(* IEC 61131-3 sources: 2026_Projet_YGO_ExcavatriceDragage/TOOLS/TEST_AUTO_CI/RESULTS/L_SIMULATION/reports (part 3) *)

(* ---- FB_Sim_PositionSensor_test.st ---- *)
(* T300 - Tests unitaires du capteur cumulatif M3. *)
TEST 'TC-T300-SEN-010 Hysteresis cumulative conserve le mot thermometre'
VAR
    fb : FB_Sim_PositionSensor;
END_VAR
    fb.Enable := TRUE;
    fb.Threshold_M := 5.0;
    fb.Hysteresis_M := 0.02;
    fb.Position_M := 4.99;
    fb();
    ASSERT_TRUE(fb.ElectricalOutput, 'Position sous seuil active DI cumulative');
    fb.Position_M := 5.01;
    fb();
    ASSERT_TRUE(fb.ElectricalOutput, 'Hysteresis maintient DI dans la bande');
    fb.Position_M := 5.03;
    fb();
    ASSERT_FALSE(fb.ElectricalOutput, 'Sortie au-dessus de seuil+hysteresis');
    fb.Position_M := 4.99;
    fb();
    ASSERT_FALSE(fb.ElectricalOutput, 'Retour dans bande ne re-declenche pas');
    fb.Position_M := 4.97;
    fb();
    ASSERT_TRUE(fb.ElectricalOutput, 'Retour sous seuil-hysteresis re-declenche');
END_TEST

TEST 'TC-T300-SEN-030 Episode intermittent est borne et rejoint la position'
VAR
    fb : FB_Sim_PositionSensor;
    i : INT;
END_VAR
    fb.Enable := TRUE;
    fb.Threshold_M := 5.0;
    fb.Position_M := 4.0;
    fb.IntermittenceActive := TRUE;
    fb.IntermittenceDurationS := 1.0;
    fb.IntermittencePeriodS := 0.12;
    fb.CycleTimeS := 0.01;
    fb();
    fb.Position_M := 6.0;
    FOR i := 1 TO 120 DO
        fb();
    END_FOR;
    ASSERT_FALSE(fb.EpisodeActive, 'Episode termine avant 1.2 s');
    ASSERT_FALSE(fb.ElectricalOutput, 'DI rejoint l etat mecanique final');
    ASSERT_GT(fb.TransitionCount, 2, 'Pertes/reprises publiees, sans front permanent');
END_TEST

TEST 'TC-T300-SEN-031 Recroisements mecaniques ne reinitialisent pas episode'
VAR
    fb : FB_Sim_PositionSensor;
    i : INT;
END_VAR
    fb.Enable := TRUE;
    fb.Threshold_M := 5.0;
    fb.Position_M := 4.0;
    fb.IntermittenceActive := TRUE;
    fb.IntermittenceDurationS := 1.0;
    fb.IntermittencePeriodS := 0.12;
    fb.CycleTimeS := 0.01;
    fb();
    FOR i := 1 TO 40 DO
        IF (i MOD 2) = 0 THEN
            fb.Position_M := 4.0;
        ELSE
            fb.Position_M := 6.0;
        END_IF;
        fb();
    END_FOR;
    fb.Position_M := 6.0;
    FOR i := 1 TO 70 DO
        fb();
    END_FOR;
    ASSERT_FALSE(fb.EpisodeActive, 'Recroisements ne prolongent pas episode au-dela de 1 s');
    ASSERT_FALSE(fb.ElectricalOutput, 'Etat final suit dernier franchissement mecanique');
END_TEST

TEST 'TC-T300-SEN-040 Cent graines deterministes bornent la stabilisation'
VAR
    fb : FB_Sim_PositionSensor;
    i : INT;
    j : INT;
END_VAR
    FOR i := 1 TO 100 DO
        fb.Enable := FALSE;
        fb();
        fb.Enable := TRUE;
        fb.Threshold_M := 5.0;
        fb.Position_M := 4.0;
        fb.IntermittenceActive := TRUE;
        fb.IntermittenceDurationS := 1.0;
        fb.IntermittencePeriodS := 0.12;
        fb.CycleTimeS := 0.01;
        fb.ScenarioSeed := DINT_TO_UDINT(i);
        fb();
        fb.Position_M := 6.0;
        FOR j := 1 TO 120 DO
            fb();
        END_FOR;
        ASSERT_FALSE(fb.EpisodeActive, 'Chaque graine termine son episode avant 1.2 s');
        ASSERT_FALSE(fb.ElectricalOutput, 'Chaque graine rejoint la position finale');
        ASSERT_GE(fb.EpisodeTogglePeriodS, 0.084, 'Periode aleatoire >= 70 % nominal');
        ASSERT_LE(fb.EpisodeTogglePeriodS, 0.156, 'Periode aleatoire <= 130 % nominal');
    END_FOR;
END_TEST

(* T300 P-A / C1-C2 — profil « BLIP COURT » : excursions electriques courtes, parametrables,
   independantes du train ~1 s ci-dessus. Signatures de la trace terrain du 2026-09-04 :
   Tremie contradictoire pendant 2 echantillons a 12,24 s ; PV reactive 1 echantillon a 14,94 s.
   Grille de test = 100 ms, celle de la trace. *)
TEST 'TC-T300-SEN-050 Blip court : largeur parametrable, deux sens, profil 1 s intact'
VAR
    fb : FB_Sim_PositionSensor;
    i : INT;
    excursions : INT;
    baseCount : UDINT;
END_VAR
    (* ---- (1) Sortie de zone, excursion 0,1 s => 1 echantillon (signature PV) ---- *)
    fb.Enable := TRUE;
    fb.Threshold_M := 5.0;
    fb.Hysteresis_M := 0.02;
    fb.CycleTimeS := 0.1;
    fb.ElectricalDelayS := 0.0;
    fb.Position_M := 4.0;
    fb();
    ASSERT_TRUE(fb.ElectricalOutput, 'Depart : dans la zone capteur');
    baseCount := fb.TransitionCount;
    fb.BlipTransitions := 1;
    fb.BlipDurationS := 0.1;
    fb.Position_M := 6.0;
    fb();
    excursions := 0;
    FOR i := 1 TO 6 DO
        fb();
        IF fb.ElectricalOutput <> fb.RawDetected THEN
            excursions := excursions + 1;
        END_IF;
    END_FOR;
    ASSERT_EQ(excursions, 1, 'Blip 0,1 s a 100 ms = 1 echantillon contradictoire');
    ASSERT_EQ(fb.TransitionCount - baseCount, 3, '1 front nominal + 2 fronts du blip');
    ASSERT_FALSE(fb.BlipActive, 'Blip borne et termine');
    ASSERT_FALSE(fb.ElectricalOutput, 'Sortie rendue a l etat mecanique final');

    (* ---- (2) Meme sens, excursion 0,2 s => 2 echantillons (signature Tremie) ---- *)
    fb.Enable := FALSE;
    fb();
    fb.Enable := TRUE;
    fb.BlipTransitions := 1;
    fb.BlipDurationS := 0.2;
    fb.Position_M := 4.0;
    fb();
    fb.Position_M := 6.0;
    fb();
    excursions := 0;
    FOR i := 1 TO 8 DO
        fb();
        IF fb.ElectricalOutput <> fb.RawDetected THEN
            excursions := excursions + 1;
        END_IF;
    END_FOR;
    ASSERT_EQ(excursions, 2, 'Blip 0,2 s a 100 ms = 2 echantillons contradictoires');
    ASSERT_FALSE(fb.ElectricalOutput, 'Sortie rendue a l etat mecanique final');

    (* ---- (3) Sens INVERSE : entree en zone (front montant) — symetrie AC5 ---- *)
    fb.Enable := FALSE;
    fb();
    fb.Enable := TRUE;
    fb.BlipTransitions := 1;
    fb.BlipDurationS := 0.2;
    fb.Position_M := 6.0;
    fb();
    ASSERT_FALSE(fb.ElectricalOutput, 'Depart : hors zone capteur');
    fb.Position_M := 4.0;
    fb();
    excursions := 0;
    FOR i := 1 TO 8 DO
        fb();
        IF fb.ElectricalOutput <> fb.RawDetected THEN
            excursions := excursions + 1;
        END_IF;
    END_FOR;
    ASSERT_EQ(excursions, 2, 'Symetrie : excursion equivalente a l entree en zone');
    ASSERT_TRUE(fb.ElectricalOutput, 'Sortie rendue a l etat mecanique final (dans la zone)');

    (* ---- (4) Blip DESACTIVE : le profil historique reste strictement inchange ---- *)
    fb.Enable := FALSE;
    fb();
    fb.Enable := TRUE;
    fb.BlipTransitions := 0;
    fb.Position_M := 4.0;
    fb();
    baseCount := fb.TransitionCount;
    fb.Position_M := 6.0;
    fb();
    excursions := 0;
    FOR i := 1 TO 10 DO
        fb();
        IF fb.ElectricalOutput <> fb.RawDetected THEN
            excursions := excursions + 1;
        END_IF;
    END_FOR;
    ASSERT_EQ(excursions, 0, 'Blip desactive : aucune excursion inventee');
    ASSERT_EQ(fb.TransitionCount - baseCount, 1, 'Blip desactive : seul le front nominal');
END_TEST

(* ---- FB_Sim_Safety_test.st ---- *)
(* =======================================================================
   Automated Unit Test - FB_Sim_Safety
   ======================================================================= *)
TEST 'TC-P13-SAF-001 Enable FALSE -> boucle AU ouverte'
VAR
    fb : FB_Sim_Safety;
END_VAR
    fb.Enable := FALSE;
    fb.SimChainOkBit := TRUE;
    fb();
    ASSERT_FALSE(fb.SimChainOk, 'Enable FALSE -> SimChainOk FALSE');
    ASSERT_FALSE(fb.SimContactorOk, 'Enable FALSE -> SimContactorOk FALSE');
END_TEST

TEST 'TC-P13-SAF-002 Pilotage boucle AU saine par SimChainOkBit et armement contacteur'
VAR
    fb : FB_Sim_Safety;
END_VAR
    fb.Enable := TRUE;
    fb.SimChainOkBit := TRUE; (* Chaine AU fermee par operateur *)
    fb();

    (* Ecoulement tempo de fermeture chaine (50ms = 60ms avancee) *)
    ADVANCE_TIME(60000000);
    fb();
    ASSERT_TRUE(fb.SimChainOk, 'SimChainOkBit TRUE -> SimChainOk TRUE apres tempo relais');

    (* Impulsion armement tenue 100ms (temps de collage contacteur) *)
    ADVANCE_TIME(10000000);
    fb.EmergencyArming := TRUE;
    fb();
    ADVANCE_TIME(110000000);
    fb();
    ASSERT_TRUE(fb.SimContactorOk, 'EmergencyArming soutenu -> SimContactorOk TRUE (engage)');

    (* Relachement impulsion -> auto-maintien *)
    ADVANCE_TIME(10000000);
    fb.EmergencyArming := FALSE;
    fb();
    ASSERT_TRUE(fb.SimContactorOk, 'Fin pulse -> Auto-maintien contacteur maintenu');
END_TEST

TEST 'TC-T306-SAF-003 Injection defaut rotation de phases par SimPhaseRotationOkBit'
VAR
    fb : FB_Sim_Safety;
END_VAR
    (* Phases saines : SimPhaseRotationOkBit=TRUE -> sortie TRUE (aucun defaut) *)
    fb.Enable := TRUE;
    fb.SimPhaseRotationOkBit := TRUE;
    fb();
    ASSERT_TRUE(fb.SimPhaseRotationOk, 'SimPhaseRotationOkBit TRUE -> SimPhaseRotationOk TRUE (phases saines)');

    (* Defaut injecte : SimPhaseRotationOkBit=FALSE -> sortie FALSE (PhaseRotationOk_DI tombe) *)
    fb.SimPhaseRotationOkBit := FALSE;
    fb();
    ASSERT_FALSE(fb.SimPhaseRotationOk, 'SimPhaseRotationOkBit FALSE -> SimPhaseRotationOk FALSE (defaut rotation de phases)');

    (* Retour a sain : nouveau passage a TRUE -> sortie TRUE *)
    fb.SimPhaseRotationOkBit := TRUE;
    fb();
    ASSERT_TRUE(fb.SimPhaseRotationOk, 'SimPhaseRotationOkBit TRUE apres FALSE -> SimPhaseRotationOk TRUE');
END_TEST

(* ---- FB_Sim_SuspendedLoad_test.st ---- *)
TEST 'TC-T300-MEC-010 Charge au repos ne cree pas d energie'
VAR
    fb : FB_Sim_SuspendedLoad;
    i : INT;
END_VAR
    fb.Enable := TRUE;
    fb.CycleTime_S := 0.01;
    FOR i := 1 TO 6000 DO
        fb();
    END_FOR;
    ASSERT_EQ(fb.Angle_Rad, 0.0, 'Angle nul sans excitation pendant 60 s');
    ASSERT_EQ(fb.AngularVelocity_RadPerS, 0.0, 'Vitesse angulaire nulle sans excitation');
END_TEST

TEST 'TC-T300-MEC-040 Acceleration excite charge et reaction reste conditionnee au frein'
VAR
    fb : FB_Sim_SuspendedLoad;
    i : INT;
END_VAR
    fb.Enable := TRUE;
    fb.CartAcceleration_Mps2 := 1.0;
    fb.BrakeMechanicallyOpen := FALSE;
    fb.CycleTime_S := 0.01;
    fb();
    ASSERT_TRUE(ABS(fb.Angle_Rad) > 0.0, 'Acceleration excite le pendule');
    ASSERT_EQ(fb.VelocityReaction_Mps, 0.0, 'Frein serre bloque reaction chariot');
    fb.BrakeMechanicallyOpen := TRUE;
    fb.CartAcceleration_Mps2 := 0.0;
    FOR i := 1 TO 10 DO
        fb();
    END_FOR;
    ASSERT_TRUE(ABS(fb.VelocityReaction_Mps) > 0.0, 'Frein ouvert publie reaction charge');
END_TEST

TEST 'TC-T300-MEC-020 Convergence pendule entre pas 10 ms et 5 ms'
VAR
    fb10 : FB_Sim_SuspendedLoad;
    fb5 : FB_Sim_SuspendedLoad;
    i : INT;
END_VAR
    fb10.Enable := TRUE;
    fb10.BrakeMechanicallyOpen := TRUE;
    fb10.CartAcceleration_Mps2 := 1.0;
    fb10.CycleTime_S := 0.01;
    fb5.Enable := TRUE;
    fb5.BrakeMechanicallyOpen := TRUE;
    fb5.CartAcceleration_Mps2 := 1.0;
    fb5.CycleTime_S := 0.005;
    fb10();
    fb5();
    fb5();
    fb10.CartAcceleration_Mps2 := 0.0;
    fb5.CartAcceleration_Mps2 := 0.0;
    FOR i := 1 TO 100 DO
        fb10();
        fb5();
        fb5();
    END_FOR;
    ASSERT_LT(ABS(fb10.Angle_Rad - fb5.Angle_Rad), 0.01,
        'Ecart angle inferieur a 10 mrad apres 1 s');
    ASSERT_LT(ABS(fb10.VelocityReaction_Mps - fb5.VelocityReaction_Mps), 0.001,
        'Ecart reaction inferieur a 1 mm/s apres 1 s');
END_TEST

(* ---- FB_Sim_Translation_test.st ---- *)
(* T300 - Tests du modele dynamique M3. *)
TEST 'TC-T300-TR-001 Etat sur desactive est P1 sans mouvement'
VAR
    fb : FB_Sim_Translation;
END_VAR
    fb.Enable := FALSE;
    fb();
    ASSERT_FALSE(fb.PosTremie, 'P1 ne doit pas annoncer Tremie');
    ASSERT_TRUE(fb.PosP1, 'Etat de repli deterministe sur P1');
    ASSERT_TRUE(fb.PosMaintenance, 'Mot thermometre P1 attendu');
    ASSERT_EQ(fb.ActualFrequency_Hz, 0.0, 'Frequence nulle');
    ASSERT_FALSE(fb.BrakeContactOpen, 'Frein ferme');
END_TEST

TEST 'TC-T300-SEN-010 Les deux extremites publient les mots thermometres valides'
VAR
    fb : FB_Sim_Translation;
    i : INT;
END_VAR
    fb.Enable := FALSE;
    fb();
    fb.Enable := TRUE;
    fb.ReqTremie := TRUE;
    fb.SpeedTgt_Pct := 100.0;
    fb.BrakeReleaseCmd := TRUE;
    fb.BrakeOpenDelayS := 0.0;
    fb.FullTravelTimeS := 0.5;
    fb.SensorElectricalDelayS := 0.0;
    FOR i := 1 TO 400 DO
        fb();
    END_FOR;
    ASSERT_TRUE(fb.PosTremie, 'Tremie active a la butee 0 m');
    ASSERT_TRUE(fb.PosPV, 'PV cumulatif actif a Tremie');
    ASSERT_TRUE(fb.PosP2, 'P2 cumulatif actif a Tremie');
    ASSERT_TRUE(fb.PosP1, 'P1 cumulatif actif a Tremie');
    ASSERT_TRUE(fb.PosMaintenance, 'Maintenance cumulatif actif a Tremie');
    ASSERT_EQ(fb.VelocityTrue_Mps, 0.0, 'Butee Tremie absorbe la vitesse chariot');

    fb.Enable := FALSE;
    fb();
    fb.Enable := TRUE;
    fb.ReqTremie := FALSE;
    fb.ReqMaintenance := TRUE;
    fb.SpeedTgt_Pct := 100.0;
    fb.BrakeReleaseCmd := TRUE;
    fb.BrakeOpenDelayS := 0.0;
    fb.FullTravelTimeS := 0.5;
    fb.SensorElectricalDelayS := 0.0;
    FOR i := 1 TO 400 DO
        fb();
    END_FOR;
    ASSERT_FALSE(fb.PosTremie, 'Tremie inactif a Maintenance');
    ASSERT_FALSE(fb.PosPV, 'PV inactif a Maintenance');
    ASSERT_FALSE(fb.PosP2, 'P2 inactif a Maintenance');
    ASSERT_FALSE(fb.PosP1, 'P1 inactif a Maintenance');
    ASSERT_FALSE(fb.PosMaintenance, 'Maintenance inactif a la butee pour mot 00000');
    ASSERT_EQ(fb.VelocityTrue_Mps, 0.0, 'Butee Maintenance absorbe la vitesse chariot');
END_TEST

TEST 'TC-T300-SEN-011 Le capteur PV commute au franchissement vers Tremie'
VAR
    fb : FB_Sim_Translation;
    i : INT;
    pvWasFalse : BOOL;
    pvTurnedTrue : BOOL;
END_VAR
    fb.Enable := TRUE;
    fb.ReqTremie := TRUE;
    fb.SpeedTgt_Pct := 100.0;
    fb.BrakeReleaseCmd := TRUE;
    fb.FullTravelTimeS := 8.0;
    fb.SensorElectricalDelayS := 0.0;
    pvWasFalse := FALSE;
    pvTurnedTrue := FALSE;
    FOR i := 1 TO 700 DO
        fb();
        IF NOT fb.PosPV THEN
            pvWasFalse := TRUE;
        END_IF;
        IF pvWasFalse AND fb.PosPV THEN
            pvTurnedTrue := TRUE;
        END_IF;
    END_FOR;
    ASSERT_TRUE(pvWasFalse, 'PV initialement inactif a P1');
    ASSERT_TRUE(pvTurnedTrue, 'PV actif apres franchissement vers Tremie');
END_TEST

TEST 'TC-T300-DRV-020 Rampe terrain 20 Hz par seconde'
VAR
    fb : FB_Sim_Translation;
    i : INT;
END_VAR
    fb.Enable := TRUE;
    fb.ReqTremie := TRUE;
    fb.SpeedTgt_Pct := 0.0;
    fb.BrakeReleaseCmd := TRUE;
    fb();
    fb.SpeedTgt_Pct := 100.0;
    FOR i := 1 TO 100 DO
        fb();
    END_FOR;
    ASSERT_GT(fb.FrequencyCmd_Hz, 19.7, 'Rampe apres 1 s >= 19.7 Hz');
    ASSERT_LT(fb.FrequencyCmd_Hz, 20.3, 'Rampe apres 1 s <= 20.3 Hz');
    ASSERT_LT(fb.ActualFrequency_Hz, fb.FrequencyCmd_Hz, 'Retour dynamique derriere la consigne');
    ASSERT_GT(fb.ActualFrequency_Hz, 16.0, 'Retour coherent avec tau 150 ms');
END_TEST

TEST 'TC-T300-BRK-025 Frein temporise et retour distinct'
VAR
    fb : FB_Sim_Translation;
    i : INT;
END_VAR
    fb.Enable := TRUE;
    fb.BrakeReleaseCmd := TRUE;
    fb.BrakeOpenDelayS := 0.10;
    fb();
    ASSERT_TRUE(fb.BrakeCoilEnergized, 'Bobine active immediatement sur ordre');
    FOR i := 1 TO 8 DO
        fb();
    END_FOR;
    ASSERT_FALSE(fb.BrakeContactOpen, 'Pas de confirmation avant 90 ms');
    fb();
    fb();
    ASSERT_TRUE(fb.BrakeMechanicallyOpen, 'Ouverture mecanique apres delai');
    ASSERT_TRUE(fb.BrakeContactOpen, 'Retour auxiliaire apres delai');
END_TEST

TEST 'TC-T300-MEC-010 Le chariot suit la frequence et excite la charge'
VAR
    fb : FB_Sim_Translation;
    i : INT;
    startPosition_M : REAL;
END_VAR
    fb.Enable := TRUE;
    fb.ReqTremie := TRUE;
    fb.SpeedTgt_Pct := 100.0;
    fb.BrakeReleaseCmd := TRUE;
    fb.BrakeOpenDelayS := 0.0;
    fb();
    startPosition_M := fb.PositionTrue_M;
    FOR i := 1 TO 100 DO
        fb();
    END_FOR;
    ASSERT_LT(fb.PositionTrue_M, startPosition_M, 'Deplacement reel vers Tremie');
    ASSERT_LT(fb.VelocityTrue_Mps, 0.0, 'Vitesse signee vers Tremie');
    ASSERT_TRUE(ABS(fb.LoadAngle_Rad) > 0.0001, 'Acceleration excite le pendule');
END_TEST

TEST 'TC-T300-MEC-030 Commandes contradictoires restent neutres'
VAR
    fb : FB_Sim_Translation;
    i : INT;
    startPosition_M : REAL;
END_VAR
    fb.Enable := TRUE;
    fb.ReqTremie := TRUE;
    fb.ReqMaintenance := TRUE;
    fb.SpeedTgt_Pct := 100.0;
    fb.BrakeReleaseCmd := TRUE;
    fb.BrakeOpenDelayS := 0.0;
    fb();
    startPosition_M := fb.PositionTrue_M;
    FOR i := 1 TO 50 DO
        fb();
    END_FOR;
    ASSERT_EQ(fb.FrequencyCmd_Hz, 0.0, 'Aucune excitation avec deux sens');
    ASSERT_EQ(fb.PositionTrue_M, startPosition_M, 'Position conservee');
END_TEST

TEST 'TC-T300-SEN-030 Episode capteur intermittent rejouable avant stabilisation'
VAR
    fb : FB_Sim_Translation;
    i : INT;
END_VAR
    fb.Enable := TRUE;
    fb.ReqMaintenance := TRUE;
    fb.SpeedTgt_Pct := 0.0;
    fb.BrakeReleaseCmd := TRUE;
    fb.BrakeOpenDelayS := 0.0;
    fb.FullTravelTimeS := 0.5;
    fb.SensorStabilizationS := 1.0;
    fb.SensorIntermittenceActive := TRUE;
    fb.SensorLoadAngleTriggerRad := 0.0;
    fb.SensorIntermittencePeriodS := 0.12;
    fb();
    fb.SpeedTgt_Pct := 100.0;
    FOR i := 1 TO 250 DO
        fb();
    END_FOR;
    ASSERT_GT(fb.SensorTransitionCount, 1, 'Au moins deux fronts DI sont publies pendant episode');
    ASSERT_FALSE(fb.PosP1, 'DI rejoint la position mecanique apres episode');
END_TEST

TEST 'TC-T300-CAM-100 Matrice 48 scenarios par 100 graines respecte invariants'
VAR
    fb : FB_Sim_Translation;
    direction : INT;
    loadProfile : INT;
    regime : INT;
    perturbation : INT;
    seed : INT;
    i : INT;
END_VAR
    FOR direction := 1 TO 2 DO
        FOR loadProfile := 1 TO 2 DO
            FOR regime := 1 TO 3 DO
                FOR perturbation := 1 TO 4 DO
                    FOR seed := 1 TO 100 DO
                        fb.Enable := FALSE;
                        fb();
                        fb.Enable := TRUE;
                        fb.ReqTremie := direction = 1;
                        fb.ReqMaintenance := direction = 2;
                        fb.SpeedTgt_Pct := 100.0;
                        fb.BrakeReleaseCmd := TRUE;
                        fb.FullTravelTimeS := 0.5;
                        fb.SensorElectricalDelayS := 0.0;
                        fb.SensorScenarioSeed := DINT_TO_UDINT(seed);
                        fb.SensorIntermittenceActive := perturbation = 3;
                        fb.SensorLoadAngleTriggerRad := 0.0;
                        IF loadProfile = 1 THEN
                            fb.LoadReactionGain_Mps2 := 0.0;
                        ELSE
                            fb.LoadReactionGain_Mps2 := 0.20;
                        END_IF;
                        IF perturbation = 4 THEN
                            fb.BrakeOpenDelayS := 0.30;
                        ELSE
                            fb.BrakeOpenDelayS := 0.0;
                        END_IF;
                        fb();
                        FOR i := 1 TO 200 DO
                            IF (regime = 2) AND (i = 80) THEN
                                fb.SpeedTgt_Pct := 0.0;
                            ELSIF (regime = 3) AND (i = 80) THEN
                                fb.SpeedTgt_Pct := 0.0;
                                fb.BrakeReleaseCmd := FALSE;
                            END_IF;
                            fb();
                            ASSERT_GE(fb.PositionTrue_M, 0.0, 'Course mecanique jamais inferieure a Tremie');
                            ASSERT_LE(fb.PositionTrue_M, 30.0, 'Course mecanique jamais superieure a Maintenance');
                            ASSERT_GE(fb.ActualFrequency_Hz, 0.0, 'Retour variateur non negatif');
                            ASSERT_LE(fb.ActualFrequency_Hz, 50.0, 'Retour variateur borne a 50 Hz');
                            IF perturbation <> 3 THEN
                                ASSERT_TRUE((NOT fb.PosTremie) OR fb.PosPV,
                                    'Mot thermometre : Tremie implique PV');
                                ASSERT_TRUE((NOT fb.PosPV) OR fb.PosP2,
                                    'Mot thermometre : PV implique P2');
                                ASSERT_TRUE((NOT fb.PosP2) OR fb.PosP1,
                                    'Mot thermometre : P2 implique P1');
                                ASSERT_TRUE((NOT fb.PosP1) OR fb.PosMaintenance,
                                    'Mot thermometre : P1 implique Maintenance');
                            END_IF;
                        END_FOR;
                    END_FOR;
                END_FOR;
            END_FOR;
        END_FOR;
    END_FOR;
END_TEST

(* T300 P-A / C4 — traversee de la faute frein dans le composite : prouve que l'entree
   descend jusqu'a FB_Sim_TranslationBrake et que la sortie remonte, sans toucher au
   nominal (premier palier d'assertions). *)
TEST 'TC-T300-BRK-041 Faute frein traverse le composite M3 (fermeture en mouvement)'
VAR
    fb : FB_Sim_Translation;
    i : INT;
END_VAR
    fb.Enable := TRUE;
    fb.ReqMaintenance := TRUE;
    fb.SpeedTgt_Pct := 100.0;
    fb.BrakeReleaseCmd := TRUE;
    fb.BrakeOpenDelayS := 0.0;
    fb();
    ASSERT_TRUE(fb.BrakeMechanicallyOpen, 'Frein ouvert au depart');
    FOR i := 1 TO 200 DO
        fb();
    END_FOR;
    ASSERT_GT(fb.ActualFrequency_Hz, 0.5, 'Chariot en mouvement (frequence non nulle)');
    ASSERT_TRUE(fb.BrakeMechanicallyOpen, 'NOMINAL : frein ouvert tant que la vitesse est non nulle');
    ASSERT_FALSE(fb.BrakeFaultCloseActive, 'Aucune faute par defaut');

    fb.BrakeFaultCloseWhileRunning := TRUE;
    FOR i := 1 TO 12 DO
        fb();
    END_FOR;
    ASSERT_TRUE(fb.BrakeFaultCloseActive, 'Faute frein relayee par le composite');
    ASSERT_GT(fb.ActualFrequency_Hz, 0.5, 'Vitesse encore non nulle a la fermeture');
    ASSERT_FALSE(fb.BrakeMechanicallyOpen, 'Faute : frein mecaniquement serre en mouvement');
END_TEST

(* T300 P-A / C3 — deceleration libre. Trace terrain 2026-09-04 : commande retiree a
   14,67 s alors que 33,98 Hz etaient retournes ; le chariot a continue d'avancer pendant
   1,49 s jusqu'a l'arret a 16,16 s. La distance de roue libre correspondante est une
   ESTIMATION (la trace ne contient aucune variable de position) : ordre de grandeur
   1,1 a 1,3 m selon la methode d'integration, jamais parcourus par le modele avant ce
   correctif qui annulait la vitesse au scan de retrait de commande.
   Le pas FullTravelTimeS est allonge (60 s) pour que le scenario reste loin des butees
   mecaniques et que l'oracle porte sur la SEULE deceleration libre, pas sur un choc. *)
TEST 'TC-T300-DRV-070 Deceleration libre : le chariot avance encore apres retrait de commande'
VAR
    fb : FB_Sim_Translation;
    i : INT;
    posAtCut_M : REAL;
END_VAR
    fb.Enable := TRUE;
    fb.ReqMaintenance := TRUE;
    fb.SpeedTgt_Pct := 100.0;
    fb.BrakeReleaseCmd := TRUE;
    fb.BrakeOpenDelayS := 0.0;
    (* Echelle par defaut du banc : palier 50 Hz (maximum variateur), 0,02 m/(Hz.s), rampe d'arret 25 Hz/s. *)
    (* Charge neutralisee : l'oracle porte sur la SEULE deceleration libre du variateur.
       Sans cela, le droop de charge (0,5 Hz par rad/s) peut faire passer ActualFrequency
       sous 39,5 Hz et rendre l'assertion de palier marginale — bruit, pas verite. *)
    fb.LoadFrequencyDroopGain_Hz := 0.0;
    fb.LoadReactionGain_Mps2 := 0.0;
    FOR i := 1 TO 400 DO
        fb();
    END_FOR;
    ASSERT_NEAR(fb.ActualFrequency_Hz, 50.0, 0.5, 'Palier 50 Hz etabli avant le retrait');
    ASSERT_LT(fb.PositionTrue_M, 30.0, 'Chariot encore hors butee (scenario non pollue)');

    (* Retrait total de la commande : plus aucune requete, consigne a zero. *)
    fb.ReqMaintenance := FALSE;
    fb.ReqTremie := FALSE;
    fb.SpeedTgt_Pct := 0.0;
    fb();
    ASSERT_GT(fb.ActualFrequency_Hz, 0.5, 'Le variateur retourne encore de la vitesse au retrait');
    posAtCut_M := fb.PositionTrue_M;

    (* Roue libre : la position doit continuer de varier tant que ActualFrequency_Hz > 0.
       Seuil = borne BASSE de la bande de reference trace (R2-O9 : 0,9 a 1,3 m). Le modele
       parcourt davantage (~2,2 m) car sa rampe de descente dure 2,0 s contre 1,49 s mesures :
       ecart de fidelite ASSUME, borne haute verifiee separement. Avant correctif : ~0,1 m. *)
    FOR i := 1 TO 300 DO
        fb();
    END_FOR;
    ASSERT_NEAR(fb.ActualFrequency_Hz, 0.0, 0.01, 'Retour variateur revenu a zero');
    ASSERT_GE(fb.PositionTrue_M - posAtCut_M, 0.9,
        'Roue libre >= borne basse trace (avant correctif : ~0,1 m)');
    ASSERT_LE(fb.PositionTrue_M - posAtCut_M, 3.0, 'Roue libre bornee (pas d emballement)');
    ASSERT_LE(fb.PositionTrue_M, 30.0, 'Course mecanique respectee');
END_TEST

(* T300 P-A / C5 — perte DEFINITIVE du capteur Tremie apres arret serre.
   Trace terrain 2026-09-04 : a 26,437 s le chariot entre en zone Tremie pendant que la
   commande est retiree ; le capteur retombe a 26,537 s et n'est JAMAIS repris sur les
   8,6 s restantes (PLAN_T300 §38 : perte unique post-arret, pas une oscillation entretenue).
   EndStopRecoilMax_M = 0 conserve le comportement historique (position ET vitesse figees,
   decision de review tracee) : les deux regimes sont verifies ici. *)
TEST 'TC-T300-SEN-052 Recul borne a la butee Tremie : DI perdue PUIS reprise oscillante (ecart trace)'
VAR
    fb : FB_Sim_Translation;
    i : INT;
    scansToFall : INT;
    scansActive : INT;
END_VAR
    (* --- (0) NON-REGRESSION : recul non autorise => comportement historique inchange --- *)
    fb.Enable := TRUE;
    fb.ReqTremie := TRUE;
    fb.SpeedTgt_Pct := 100.0;
    fb.BrakeReleaseCmd := TRUE;
    fb.BrakeOpenDelayS := 0.0;
    fb.SensorElectricalDelayS := 0.0;
    fb.EndStopRecoilMax_M := 0.0;
    (* T361 — pas de temps PINCE ici : l'oracle de ce cas est le recul a la butee, pas
       l'echelle odometrique. Le scenario vient de la trace du 2026-09-04 (quelques
       secondes de trajet) et le defaut du FB est passe de 8,0 s a 37,5 s pour s'aligner
       sur le gain reel : sans ce pas explicite, 900 scans (9 s) ne suffiraient plus a
       atteindre la butee Tremie depuis 20 m et le cas testerait autre chose que son objet. *)
    fb.FullTravelTimeS := 8.0;
    FOR i := 1 TO 900 DO
        fb();
    END_FOR;
    ASSERT_TRUE(fb.PosTremie, 'Historique : DI Tremie TENUE a la butee quand le recul est interdit');
    ASSERT_NEAR(fb.PositionTrue_M, 0.0, 0.001, 'Historique : position figee a la butee');

    (* --- (1) Recul borne autorise : la charge ressort le chariot de la zone --- *)
    fb.Enable := FALSE;
    fb();
    fb.Enable := TRUE;
    fb.EndStopRecoilMax_M := 0.5;
    fb.LoadReactionGain_Mps2 := 2.0;
    FOR i := 1 TO 900 DO
        fb();
    END_FOR;
    ASSERT_TRUE(fb.PosTremie, 'PRECONDITION : zone Tremie atteinte (recul = 0,5 m autorise)');

    (* Commande retiree a l'instant de l' entree en zone (sequence exacte de la trace). *)
    fb.ReqTremie := FALSE;
    fb.SpeedTgt_Pct := 0.0;
    scansToFall := 0;
    FOR i := 1 TO 600 DO
        fb();
        IF (NOT fb.PosTremie) AND (scansToFall = 0) THEN
            scansToFall := i;
        END_IF;
    END_FOR;
    ASSERT_GT(scansToFall, 0, 'DI Tremie RETOMBE apres l arret serre (recul borne)');
    (* Boucle a 600 scans, seuil a 300 : assertion NON tautologique, marge reelle au-dessus
       de la valeur mesuree (256 scans). *)
    ASSERT_LE(scansToFall, 300, 'Perte dans un temps borne (<= 3 s a 10 ms)');

    (* Perte DURABLE : le capteur ne se reactive pas de facon entretenue ensuite. *)
    scansActive := 0;
    FOR i := 1 TO 500 DO
        fb();
        IF fb.PosTremie THEN
            scansActive := scansActive + 1;
        END_IF;
    END_FOR;
    (* ⚠️ LIMITE CONNUE — NON MASQUEE. Le modele reduit n'a AUCUNE friction de chariot ni
       raideur de cable : le pendule amorti ramene le chariot dans la zone capteur par
       oscillations. La perte est donc BORNEE, mais pas encore DEFINITIVE comme sur la trace
       terrain (PLAN_T300 §38 : « perte unique post-arret, pas une oscillation entretenue »).
       Fermer cet ecart exige un parametre physique nouveau (friction de roulement / raideur
       de cable), hors perimetre de ce lot et non calibrable sans mesure terrain : ce test
       CARACTERISE l'etat reel, il ne le valide pas. Mesure : 106 scans actifs sur 500
       (21 %), contre 0 attendu par la trace. Assertion volontairement en enveloppe. *)
    ASSERT_LE(scansActive, 150, 'Perte BORNEE mais NON DEFINITIVE : ecart trace documente');
END_TEST

(* =========================================================================
   T361 VOLET A — ALIGNEMENT DU RATIO ODOMETRIQUE BANC / ESTIMATEUR
   =========================================================================
   Le banc et l'estimateur integrent la MEME frequence retournee, mais avec deux
   echelles construites separement :
     - estimateur (CODE/I_TRANSLATION/FB_Translation_PositionEstimator.st:153/155) :
       dx = f x GainMetersPerHzSec x dt, gain cable en PRG_05_Translation.st:591 sur
       GVL_PERSISTENT._TranslationGainMetersPerHzSec = 0,02 m/(Hz.s) (1 m/s a 50 Hz) ;
     - banc (ce FB) : dx = f x (CST_PositionAtMaintenance / (40 x FullTravelTimeS)) x dt.
   Tant que les deux echelles divergent, la position estimee prend un retard constant et
   CHAQUE franchissement de capteur produit un saut de recalage — c'est exactement ce que
   montre la trace Suivi_74 (sauts de 4,53 / 9,12 / 4,59 m, AUDIT_T360). Avec l'echelle
   historique 8,0 s le rapport valait 0,09375 / 0,02 = 4,7.
   Les deux cas ci-dessous comparent le banc a l'expression EXACTE de l'estimateur :
   ils echouent si l'une des deux echelles bouge sans l'autre. *)

TEST 'TC-T361-ALIGN-001 Ratio odometrique du banc = gain reel 0,02 m/(Hz.s)'
VAR
    fb : FB_Sim_Translation;
    i : INT;
END_VAR
    fb.Enable := TRUE;
    fb.ReqMaintenance := TRUE;
    fb.SpeedTgt_Pct := 100.0;
    fb.BrakeReleaseCmd := TRUE;
    fb.BrakeOpenDelayS := 0.0;
    (* Charge neutralisee : l'oracle porte sur l'ECHELLE seule, pas sur la reaction du pendule. *)
    fb.LoadReactionGain_Mps2 := 0.0;
    FOR i := 1 TO 400 DO
        fb();
    END_FOR;
    ASSERT_NEAR(fb.ActualFrequency_Hz, 50.0, 0.5, 'Palier 50 Hz (maximum variateur) etabli avant lecture du ratio');
    ASSERT_NEAR(fb.VelocityTrue_Mps / fb.ActualFrequency_Hz, 0.02, 0.0002,
        'Ratio banc (m/s par Hz) = _TranslationGainMetersPerHzSec (ancien : 0,09375)');
END_TEST

TEST 'TC-T361-ALIGN-002 Distance banc = integrale f x 0,02 m/(Hz.s) sur 6 s'
VAR
    fb : FB_Sim_Translation;
    i : INT;
    posStart_M : REAL;
    integralHzS : REAL;
END_VAR
    fb.Enable := TRUE;
    fb.ReqTremie := TRUE;
    fb.SpeedTgt_Pct := 100.0;
    fb.BrakeReleaseCmd := TRUE;
    fb.BrakeOpenDelayS := 0.0;
    fb.SensorElectricalDelayS := 0.0;
    fb.LoadReactionGain_Mps2 := 0.0;
    (* 2 s pour etablir le palier, puis 6 s de mesure (600 scans a 10 ms) largement
       a l'ecart des butees : 20 m -> ~15,2 m a 0,8 m/s. *)
    FOR i := 1 TO 200 DO
        fb();
    END_FOR;
    posStart_M := fb.PositionTrue_M;
    integralHzS := 0.0;
    FOR i := 1 TO 600 DO
        fb();
        integralHzS := integralHzS + fb.ActualFrequency_Hz * 0.010;
    END_FOR;
    (* Tolerance 0,25 m (soit ~5 % de 4,8 m) : elle couvre la seule trainee de 1er ordre du
       modele de vitesse, pas une erreur d'echelle — un ecart d'echelle de 4,7 ferait
       diverger les deux membres de plusieurs metres. *)
    ASSERT_NEAR(posStart_M - fb.PositionTrue_M, integralHzS * 0.02, 0.25,
        'Distance parcourue par le banc = position reconstituee par l estimateur odometrique');
END_TEST

(* Echelle de la consigne : PRG_02 envoie SpeedCmd_Pct = f / 50 Hz x 100.
   20 Hz d'approche reels = 40 % doivent redonner 20 Hz (pas 16 Hz). Charge neutralisee. *)
TEST 'TC-T417-SCALE-001 Consigne 40 pct = 20 Hz et 100 pct = 50 Hz'
VAR
    fbApproach : FB_Sim_Translation;
    fbMax : FB_Sim_Translation;
    i : INT;
END_VAR
    fbApproach.Enable := TRUE;
    fbApproach.ReqMaintenance := TRUE;
    fbApproach.SpeedTgt_Pct := 40.0;
    fbApproach.BrakeReleaseCmd := TRUE;
    fbApproach.BrakeOpenDelayS := 0.0;
    fbApproach.LoadFrequencyDroopGain_Hz := 0.0;
    fbApproach.LoadReactionGain_Mps2 := 0.0;
    fbMax.Enable := TRUE;
    fbMax.ReqMaintenance := TRUE;
    fbMax.SpeedTgt_Pct := 100.0;
    fbMax.BrakeReleaseCmd := TRUE;
    fbMax.BrakeOpenDelayS := 0.0;
    fbMax.LoadFrequencyDroopGain_Hz := 0.0;
    fbMax.LoadReactionGain_Mps2 := 0.0;
    FOR i := 1 TO 400 DO
        fbApproach();
        fbMax();
    END_FOR;
    ASSERT_NEAR(fbApproach.ActualFrequency_Hz, 20.0, 0.05, '40 pct de 50 Hz = 20 Hz en regime etabli');
    ASSERT_NEAR(fbMax.ActualFrequency_Hz, 50.0, 0.05, '100 pct = 50 Hz (maximum variateur)');
END_TEST

(* Rampe d'arret : trace reelle ~25 Hz/s (rampe variateur). Pente mesuree sur la fenetre
   utile 10 Hz -> ~4 Hz, apres le transitoire du filtre de 1er ordre. Charge neutralisee. *)
TEST 'TC-T417-DECEL-001 Pente d arret 25 Hz/s depuis l approche 20 Hz'
VAR
    fb : FB_Sim_Translation;
    i : INT;
    f1_Hz : REAL;
END_VAR
    fb.Enable := TRUE;
    fb.ReqMaintenance := TRUE;
    fb.SpeedTgt_Pct := 40.0;
    fb.BrakeReleaseCmd := TRUE;
    fb.BrakeOpenDelayS := 0.0;
    fb.LoadFrequencyDroopGain_Hz := 0.0;
    fb.LoadReactionGain_Mps2 := 0.0;
    FOR i := 1 TO 400 DO
        fb();
    END_FOR;
    ASSERT_NEAR(fb.ActualFrequency_Hz, 20.0, 0.05, 'Approche 20 Hz etablie avant le retrait');
    fb.SpeedTgt_Pct := 0.0;
    i := 0;
    WHILE (fb.ActualFrequency_Hz > 10.0) AND (i < 300) DO
        fb();
        i := i + 1;
    END_WHILE;
    f1_Hz := fb.ActualFrequency_Hz;
    FOR i := 1 TO 20 DO
        fb();
    END_FOR;
    ASSERT_NEAR((f1_Hz - fb.ActualFrequency_Hz) / 0.2, 25.0, 1.0, 'Pente de decroissance = 25 Hz/s');
END_TEST

(* Depassement apres retrait de commande a l'approche : ordre de grandeur de la trace reelle
   (~0,25 m, gain 0,02 m/(Hz.s) provisoire). Bande large : cible a confirmer par la trace 10 ms. *)
TEST 'TC-T417-OVERSHOOT-001 Depassement apres retrait a 20 Hz'
VAR
    fb : FB_Sim_Translation;
    i : INT;
    posAtCut_M : REAL;
    overshoot_M : REAL;
END_VAR
    fb.Enable := TRUE;
    fb.ReqMaintenance := TRUE;
    fb.SpeedTgt_Pct := 40.0;
    fb.BrakeReleaseCmd := TRUE;
    fb.BrakeOpenDelayS := 0.0;
    fb.LoadFrequencyDroopGain_Hz := 0.0;
    fb.LoadReactionGain_Mps2 := 0.0;
    FOR i := 1 TO 400 DO
        fb();
    END_FOR;
    ASSERT_NEAR(fb.ActualFrequency_Hz, 20.0, 0.05, 'Approche 20 Hz etablie avant le retrait');
    fb.ReqMaintenance := FALSE;
    fb.SpeedTgt_Pct := 0.0;
    fb();
    posAtCut_M := fb.PositionTrue_M;
    FOR i := 1 TO 300 DO
        fb();
    END_FOR;
    overshoot_M := fb.PositionTrue_M - posAtCut_M;
    ASSERT_GE(overshoot_M, 0.15, 'Depassement >= 0,15 m (ordre de grandeur trace reelle)');
    ASSERT_LE(overshoot_M, 0.35, 'Depassement <= 0,35 m (ordre de grandeur trace reelle)');
END_TEST

(* Acceleration du banc : chariot ET frequence retournee x facteur. L'estimateur reel integre
   f_retournee x 0,02 : il doit retrouver la distance du chariot (aucun saut de recalage). *)
TEST 'TC-SIMSPEED-001 Facteur 3 : chariot 3 m/s a 50 Hz et distance = integrale f retournee x 0,02'
VAR
    fb : FB_Sim_Translation;
    i : INT;
    posStart_M : REAL;
    integralHzS : REAL;
END_VAR
    fb.Enable := TRUE;
    fb.ReqTremie := TRUE;
    fb.SpeedTgt_Pct := 100.0;
    fb.SpeedFactor := 3.0;
    fb.BrakeReleaseCmd := TRUE;
    fb.BrakeOpenDelayS := 0.0;
    fb.SensorElectricalDelayS := 0.0;
    fb.LoadReactionGain_Mps2 := 0.0;
    FOR i := 1 TO 300 DO
        fb();
    END_FOR;
    ASSERT_NEAR(fb.ActualFrequency_Hz, 150.0, 3.0, 'frequence retournee = 3 x 50 Hz');
    ASSERT_NEAR(fb.VelocityTrue_Mps, -3.0, 0.15, 'chariot a 3 m/s (1 m/s reel x 3)');
    posStart_M := fb.PositionTrue_M;
    integralHzS := 0.0;
    FOR i := 1 TO 200 DO
        fb();
        integralHzS := integralHzS + fb.ActualFrequency_Hz * 0.010;
    END_FOR;
    ASSERT_NEAR(posStart_M - fb.PositionTrue_M, integralHzS * 0.02, 0.25,
        'estimation (f retournee x 0,02) = distance du chariot : aucun saut de recalage');
END_TEST

TEST 'TC-SIMSPEED-002 Facteur borne a 5, facteur < 1 ramene a 1'
VAR
    fb : FB_Sim_Translation;
    fbLow : FB_Sim_Translation;
    i : INT;
END_VAR
    fb.Enable := TRUE;
    fb.ReqTremie := TRUE;
    fb.SpeedTgt_Pct := 100.0;
    fb.SpeedFactor := 10.0;
    fb.BrakeReleaseCmd := TRUE;
    fb.BrakeOpenDelayS := 0.0;
    fb.LoadReactionGain_Mps2 := 0.0;
    fbLow.Enable := TRUE;
    fbLow.ReqTremie := TRUE;
    fbLow.SpeedTgt_Pct := 100.0;
    fbLow.SpeedFactor := 0.0;
    fbLow.BrakeReleaseCmd := TRUE;
    fbLow.BrakeOpenDelayS := 0.0;
    fbLow.LoadReactionGain_Mps2 := 0.0;
    FOR i := 1 TO 300 DO
        fb();
        fbLow();
    END_FOR;
    ASSERT_NEAR(fb.ActualFrequency_Hz, 250.0, 5.0, 'facteur 10 borne a 5 : 250 Hz retournes');
    ASSERT_NEAR(fbLow.ActualFrequency_Hz, 50.0, 1.0, 'facteur 0 ramene a 1 : 50 Hz retournes');
    ASSERT_NEAR(fbLow.VelocityTrue_Mps, -1.0, 0.05, 'facteur 1 : 1 m/s reel a 50 Hz');
END_TEST

(* ---- FB_Sim_TranslationBrake_test.st ---- *)
TEST 'TC-T300-BRK-010 Bobine mecanique et contact restent distincts'
VAR
    fb : FB_Sim_TranslationBrake;
    i : INT;
END_VAR
    fb.Enable := TRUE;
    fb.ReleaseCmd := TRUE;
    fb.OpenDelay_S := 0.10;
    fb.ContactDelay_S := 0.01;
    fb.CycleTime_S := 0.01;
    FOR i := 1 TO 9 DO
        fb();
    END_FOR;
    ASSERT_TRUE(fb.CoilEnergized, 'Bobine immediate');
    ASSERT_FALSE(fb.MechanicallyOpen, 'Effet mecanique pas avant delai');
    fb();
    fb();
    ASSERT_TRUE(fb.MechanicallyOpen, 'Ouverture mecanique apres 100 ms');
    fb();
    ASSERT_TRUE(fb.ContactOpen, 'Contact apres effet mecanique');
END_TEST

TEST 'TC-T300-BRK-020 Serrage attend vitesse nulle'
VAR
    fb : FB_Sim_TranslationBrake;
    i : INT;
END_VAR
    fb.Enable := TRUE;
    fb.ReleaseCmd := TRUE;
    fb.OpenDelay_S := 0.0;
    fb.CycleTime_S := 0.01;
    fb();
    fb.ReleaseCmd := FALSE;
    fb.ActualFrequency_Hz := 2.0;
    FOR i := 1 TO 20 DO
        fb();
    END_FOR;
    ASSERT_TRUE(fb.MechanicallyOpen, 'Frein reste ouvert tant que vitesse non nulle');
    fb.ActualFrequency_Hz := 0.0;
    FOR i := 1 TO 10 DO
        fb();
    END_FOR;
    ASSERT_FALSE(fb.MechanicallyOpen, 'Frein serre apres 90 ms a vitesse nulle');
END_TEST

(* T300 P-A / C4 — rejeu EXACT du defaut terrain du 2026-09-04 (trace M3, 26,437 s) :
   contact frein ferme alors que le variateur retourne encore 10,00 Hz (State.ErrorId=64).
   La branche de FAUTE est explicite et le defaut de l'entree est FALSE : le chemin nominal
   reste celui de TC-T300-BRK-020, dont la garde 0,5 Hz est validee par la MEME trace
   (frein ouvert a 0,60 Hz a 16,04 s, ferme a 0,00 Hz a 16,16 s). *)
TEST 'TC-T300-BRK-040 Faute explicite : frein M3 se ferme a 10 Hz (rejeu trace 26,437 s)'
VAR
    fb : FB_Sim_TranslationBrake;
    i : INT;
END_VAR
    fb.Enable := TRUE;
    fb.ReleaseCmd := TRUE;
    fb.OpenDelay_S := 0.0;
    fb.CloseDelay_S := 0.09;
    fb.ContactDelay_S := 0.01;
    fb.CycleTime_S := 0.01;
    fb();
    ASSERT_TRUE(fb.MechanicallyOpen, 'Frein ouvert par la commande de desserrage');
    ASSERT_FALSE(fb.FaultCloseActive, 'Faute inactive par defaut');

    (* Scenario terrain : commande retiree ET variateur retournant encore 10,00 Hz. *)
    fb.ReleaseCmd := FALSE;
    fb.ActualFrequency_Hz := 10.0;
    FOR i := 1 TO 20 DO
        fb();
    END_FOR;
    ASSERT_FALSE(fb.FaultCloseActive, 'Aucune faute injectee');
    ASSERT_TRUE(fb.MechanicallyOpen, 'NOMINAL conserve : frein OUVERT a 10,00 Hz (garde 0,5 Hz)');
    ASSERT_TRUE(fb.ContactOpen, 'NOMINAL conserve : contact toujours ouvert a 10,00 Hz');

    (* Injection explicite : fermeture hors vitesse nulle, APRES le delai de faute.
       Oracle discriminateur : si le delai de faute etait ignore, la faute serait appliquee
       des le 1er scan et l'assertion ci-dessous echouerait. *)
    fb.FaultCloseWhileRunning := TRUE;
    fb.FaultCloseDelay_S := 0.5;
    FOR i := 1 TO 4 DO
        fb();
    END_FOR;
    ASSERT_FALSE(fb.FaultCloseActive, 'Faute NON appliquee avant FaultCloseDelay_S');
    ASSERT_TRUE(fb.MechanicallyOpen, 'Frein encore ouvert pendant le delai de faute');
    FOR i := 1 TO 60 DO
        fb();
    END_FOR;
    ASSERT_TRUE(fb.FaultCloseActive, 'Branche de faute appliquee apres le delai');
    ASSERT_FALSE(fb.CoilEnergized, 'Faute : bobine retombee (etat electrique coherent)');
    ASSERT_FALSE(fb.MechanicallyOpen, 'Faute : frein MECANIQUEMENT serre a 10,00 Hz');
    ASSERT_FALSE(fb.ContactOpen, 'Faute : contact frein ferme publie a 10,00 Hz');

    (* Retrait du stimulus : retour au chemin nominal, sans etat residuel. *)
    fb.FaultCloseWhileRunning := FALSE;
    fb();
    ASSERT_FALSE(fb.FaultCloseActive, 'Retrait du stimulus : faute retombee');
END_TEST

(* ---- FB_Sim_TranslationDrive_test.st ---- *)
TEST 'TC-T300-DRV-010 Drive rampe et reponse premier ordre'
VAR
    fb : FB_Sim_TranslationDrive;
    i : INT;
END_VAR
    fb.Enable := TRUE;
    fb.FrequencyTgt_Hz := 40.0;
    fb.CycleTime_S := 0.01;
    FOR i := 1 TO 100 DO
        fb();
    END_FOR;
    ASSERT_GT(fb.FrequencyCmd_Hz, 19.7, 'Rampe 20 Hz/s apres 1 s');
    ASSERT_LT(fb.FrequencyCmd_Hz, 20.3, 'Rampe bornee apres 1 s');
    ASSERT_LT(fb.ActualFrequency_Hz, fb.FrequencyCmd_Hz, 'Retour derriere la consigne');
    ASSERT_TRUE(fb.Ready, 'Brique prete sous Enable');
END_TEST

TEST 'TC-T300-DRV-030 Charge reduit retour sans inverser la frequence'
VAR
    fb : FB_Sim_TranslationDrive;
    i : INT;
    unloaded_Hz : REAL;
END_VAR
    fb.Enable := TRUE;
    fb.FrequencyTgt_Hz := 40.0;
    fb.CycleTime_S := 0.01;
    FOR i := 1 TO 300 DO
        fb();
    END_FOR;
    unloaded_Hz := fb.ActualFrequency_Hz;
    fb.LoadAngularVelocity_RadPerS := 8.0;
    fb();
    ASSERT_LT(fb.ActualFrequency_Hz, unloaded_Hz, 'Droop charge visible au PDO');
    ASSERT_GE(fb.ActualFrequency_Hz, 0.0, 'Frequence jamais negative');
END_TEST

TEST 'TC-T300-DRV-050 Pas de 100 ms conserve le temps physique'
VAR
    fb : FB_Sim_TranslationDrive;
END_VAR
    fb.Enable := TRUE;
    fb.FrequencyTgt_Hz := 40.0;
    fb.AccelRate_HzPerS := 20.0;
    fb.CycleTime_S := 0.100;
    fb();
    ASSERT_NEAR(fb.FrequencyCmd_Hz, 2.0, 0.001,
        'A 100 ms, la rampe 20 Hz/s avance de 2 Hz');
    fb();
    ASSERT_NEAR(fb.FrequencyCmd_Hz, 4.0, 0.001,
        'Le deuxieme cycle conserve la meme duree physique');
END_TEST

(* ---- FB_SimBench_test.st ---- *)
SETUP
VAR
    FB_Bench : FB_SimBench;
    FB_SimEnc : FB_Sim_Encoder;
    FB_SimJoy : FB_Sim_Joystick;
    FB_SimSafe : FB_Sim_Safety;
    FB_SimTrans : FB_Sim_Translation;
    RawPosM1 : UDINT := 0;
    RawPosM2 : UDINT := 0;
END_VAR
END_SETUP

TEST 'TC-P03-001 Dynamique Enable : neutralisation initiale, transition Ready au repos, puis coupure'
    (* Scan 0 : Enable=FALSE -> Neutralisation *)
    FB_Bench(Enable := FALSE, RawPosM1 := RawPosM1, RawPosM2 := RawPosM2);
    ASSERT_FALSE(FB_Bench.Ready, 'Enable=FALSE -> Ready=FALSE (neutralise)');

    ADVANCE_TIME(10000000);

    (* Scan 1 : Enable=TRUE -> SimBench actif *)
    FB_Bench(Enable := TRUE, RawPosM1 := RawPosM1, RawPosM2 := RawPosM2);
    ASSERT_TRUE(FB_Bench.Ready, 'Enable=TRUE -> Ready=TRUE (nominal)');

    ADVANCE_TIME(10000000);

    (* Scan 2 : Enable=FALSE -> Re-neutralisation *)
    FB_Bench(Enable := FALSE, RawPosM1 := RawPosM1, RawPosM2 := RawPosM2);
    ASSERT_FALSE(FB_Bench.Ready, 'Coupure -> Ready retombe a FALSE');
END_TEST

TEST 'TC-P13-001 Sim_Safety : neutralisation sans Enable'
    FB_SimSafe(Enable := FALSE);
    ASSERT_FALSE(FB_SimSafe.SimChainOk, 'AU non ferme');
    ASSERT_FALSE(FB_SimSafe.SimContactorOk, 'Contacteur coupe');
END_TEST

(* =========================================================================
   AF-13 — FB_SimBench (TC-P13-010/011/012/013)
   ========================================================================= *)

TEST 'TC-P13-010 SimBench Enable=FALSE neutralise tout le banc'
    FB_Bench(Enable := FALSE, RawPosM1 := RawPosM1, RawPosM2 := RawPosM2);
    ASSERT_FALSE(FB_Bench.Ready, 'Enable=FALSE -> Ready=FALSE');
    ASSERT_FALSE(FB_Bench.Busy, 'Enable=FALSE -> Busy=FALSE');
    ASSERT_FALSE(FB_Bench.Done, 'Enable=FALSE -> Done=FALSE');
END_TEST

(* =========================================================================
   T342 — CR2 : reinjection silencieuse du comptage brut (RawPosM2 = 0 -> 1 100 000 pts)
   Remplace TC-P13-014 « initialise les codeurs absolus vierges » (ID par ailleurs porte
   par l'AF-13 pour le capteur haut TOP : collision d'ID levee au passage) : le banc
   n'initialise PLUS rien, le cas « memoire vierge » est couvert par l'initialisation
   declaree GVL_PERSISTENT._SimEncoderRawPosM1/M2 := 1000000.
   ========================================================================= *)

TEST 'TC-T342-010 AUCUNE reinjection du comptage brut : un 0 reel du codeur est conserve (pas de saut post-AU)'
    (* Etat EXACT de l'incident T338 (saut 8,50 -> 204,677 m apres reactivation du banc) :
       memoire codeur a 0, banc desactive (Enable=FALSE), puis reactivation du banc
       (GVL_Simulation.SimulationModeActive FALSE -> TRUE). Le comptage brut est un entier
       SIGNE dont le zero est arbitraire (correctif T338) : le banc ne doit JAMAIS y
       substituer une origine device, sous peine d'une teleportation de
       1 100 000 pts / 4096 pts/m = 268,55 m sur la position publiee, sans mouvement
       ni defaut, reference de homing conservee. *)
    FB_Bench(Enable := FALSE, RawPosM1 := RawPosM1, RawPosM2 := RawPosM2);
    RawPosM1 := 0;
    RawPosM2 := 0;
    ADVANCE_TIME(10000000);
    FB_Bench(Enable := TRUE, RawPosM1 := RawPosM1, RawPosM2 := RawPosM2);
    ASSERT_EQ(RawPosM2, 0, 'Reactivation : la memoire codeur M2 reste a 0 (aucune reinjection du banc)');
    ASSERT_EQ(FB_Bench.Winch.COD2_PosValue, 0, 'Aucun saut publie sur COD2_PosValue (268,55 m si reinjecte)');
    ASSERT_EQ(RawPosM1, 0, 'Reactivation : la memoire codeur M1 reste a 0 (aucune reinjection du banc)');
    ASSERT_EQ(FB_Bench.Winch.COD1_PosValue, 0, 'Aucun saut publie sur COD1_PosValue');
END_TEST

TEST 'TC-T342-011 Reactivation du banc : le comptage brut conserve sa valeur courante (aucune ecriture du banc)'
    (* Non-regression du meme invariant sur une memoire MID-COURSE (296 459 pts = la valeur
       R0 reconstituee par le diagnostic T338) : quelle que soit la valeur, la reactivation
       ne produit aucun ecart, et le banc reste sans ecriture sur la memoire du codeur. *)
    FB_Bench(Enable := FALSE, RawPosM1 := RawPosM1, RawPosM2 := RawPosM2);
    RawPosM1 := 296459;
    RawPosM2 := 296459;
    ADVANCE_TIME(10000000);
    FB_Bench(Enable := TRUE, RawPosM1 := RawPosM1, RawPosM2 := RawPosM2);
    ASSERT_EQ(RawPosM2, 296459, 'Memoire M2 mid-course inchangee par la reactivation du banc');
    ASSERT_EQ(FB_Bench.Winch.COD2_PosValue, 296459, 'Position publiee = comptage brut, sans ecart');
    ASSERT_EQ(RawPosM1, 296459, 'Memoire M1 mid-course inchangee par la reactivation du banc');
    ASSERT_EQ(FB_Bench.Winch.COD1_PosValue, 296459, 'Position publiee = comptage brut, sans ecart');
END_TEST

TEST 'TC-P13-011 SimBench 0 lecture GVL en interne (essai manuel — stub)'
    (* Stub : TC-P13-011 verifie que FB_SimBench ne lit aucune variable GVL_* en interne
       (toutes les entrees passees en parametres par PRG_02_Acquisition). Verification
       statique de code, non automatisable en boite noire. (essai manuel — stub) *)
    ASSERT_TRUE(TRUE, 'Stub : verification statique 0 lecture GVL (essai manuel)');
END_TEST

TEST 'TC-P13-012 SimBench polarite frein M1 : M1_BrakeIsOpen_DI := M1_BrakeCmd'
    FB_Bench(Enable := TRUE, M1_BrakeCmd := TRUE, RawPosM1 := RawPosM1, RawPosM2 := RawPosM2);
    ASSERT_TRUE(FB_Bench.Winch.M1_BrakeIsOpen_DI, 'M1_BrakeCmd=TRUE -> M1_BrakeIsOpen_DI=TRUE (jamais NOT)');
    ADVANCE_TIME(10000000);
    FB_Bench(Enable := TRUE, M1_BrakeCmd := FALSE, RawPosM1 := RawPosM1, RawPosM2 := RawPosM2);
    ASSERT_FALSE(FB_Bench.Winch.M1_BrakeIsOpen_DI, 'M1_BrakeCmd=FALSE -> M1_BrakeIsOpen_DI=FALSE');
END_TEST

TEST 'TC-T318-010 SimBench cable nominal independent du Kobold et injection explicite'
    FB_Bench(Enable := TRUE, SimKoboldContactValue := TRUE,
             SimM2TensionedCableFaultInject := FALSE,
             RawPosM1 := RawPosM1, RawPosM2 := RawPosM2);
    ASSERT_TRUE(FB_Bench.Winch.M2_TensionedCable_DI,
                'Kobold ne produit pas de mou de cable sans injection explicite');
    FB_Bench(Enable := TRUE, SimM2TensionedCableFaultInject := TRUE,
             RawPosM1 := RawPosM1, RawPosM2 := RawPosM2);
    ASSERT_FALSE(FB_Bench.Winch.M2_TensionedCable_DI,
                 'Injection explicite -> cable non tendu');
END_TEST

TEST 'TC-T318-020 Diagnostic electrique desactive publie etat neutre'
    FB_Bench(Enable := TRUE, SimWinchElectricalDiagnosticsActive := FALSE,
             RawPosM1 := RawPosM1, RawPosM2 := RawPosM2);
    ASSERT_EQ(FB_Bench.MotorTorqueM1_Nm, 0.0, 'Diagnostic M1 OFF -> couple neutre');
    ASSERT_FALSE(FB_Bench.MotorIsStalledM1, 'Diagnostic M1 OFF -> stall FALSE');
    ASSERT_EQ(FB_Bench.MotorTorqueM2_Nm, 0.0, 'Diagnostic M2 OFF -> couple neutre');
    ASSERT_FALSE(FB_Bench.MotorIsStalledM2, 'Diagnostic M2 OFF -> stall FALSE');
END_TEST

TEST 'TC-P13-015 SimBench delai frein M1 opt-in (T316) : SimWinchBrakeOpenDelayS retarde M1_BrakeIsOpen_DI sans jamais inverser la polarite'
    (* Delai desactive (0.0) : comportement historique, bascule au meme scan *)
    FB_Bench(Enable := TRUE, M1_BrakeCmd := TRUE, SimWinchBrakeOpenDelayS := 0.0, RawPosM1 := RawPosM1, RawPosM2 := RawPosM2);
    ASSERT_TRUE(FB_Bench.Winch.M1_BrakeIsOpen_DI, 'Delai=0.0 -> ouverture instantanee (non-regression)');
    ADVANCE_TIME(10000000);
    FB_Bench(Enable := TRUE, M1_BrakeCmd := FALSE, SimWinchBrakeOpenDelayS := 0.0, RawPosM1 := RawPosM1, RawPosM2 := RawPosM2);
    ASSERT_FALSE(FB_Bench.Winch.M1_BrakeIsOpen_DI, 'Retour delai=0.0 avant test delai>0 : etat repos');

    (* Delai actif (50 ms = 5 scans a 10 ms) : la DI reste fausse pendant le delai puis bascule *)
    ADVANCE_TIME(10000000);
    FB_Bench(Enable := TRUE, M1_BrakeCmd := TRUE, SimWinchDynamicsActive := TRUE, SimWinchBrakeOpenDelayS := 0.042, RawPosM1 := RawPosM1, RawPosM2 := RawPosM2);
    ASSERT_FALSE(FB_Bench.Winch.M1_BrakeIsOpen_DI, 'Scan 1/5 du delai : M1_BrakeIsOpen_DI reste FALSE, jamais TRUE en avance');
    ADVANCE_TIME(10000000);
    FB_Bench(Enable := TRUE, M1_BrakeCmd := TRUE, SimWinchDynamicsActive := TRUE, SimWinchBrakeOpenDelayS := 0.042, RawPosM1 := RawPosM1, RawPosM2 := RawPosM2);
    ASSERT_FALSE(FB_Bench.Winch.M1_BrakeIsOpen_DI, 'Scan 2/5 du delai : toujours FALSE');
    ADVANCE_TIME(10000000);
    FB_Bench(Enable := TRUE, M1_BrakeCmd := TRUE, SimWinchDynamicsActive := TRUE, SimWinchBrakeOpenDelayS := 0.042, RawPosM1 := RawPosM1, RawPosM2 := RawPosM2);
    ASSERT_FALSE(FB_Bench.Winch.M1_BrakeIsOpen_DI, 'Scan 3/5 du delai : toujours FALSE');
    ADVANCE_TIME(10000000);
    FB_Bench(Enable := TRUE, M1_BrakeCmd := TRUE, SimWinchDynamicsActive := TRUE, SimWinchBrakeOpenDelayS := 0.042, RawPosM1 := RawPosM1, RawPosM2 := RawPosM2);
    ASSERT_FALSE(FB_Bench.Winch.M1_BrakeIsOpen_DI, 'Scan 4/5 du delai : toujours FALSE');
    ADVANCE_TIME(10000000);
    FB_Bench(Enable := TRUE, M1_BrakeCmd := TRUE, SimWinchDynamicsActive := TRUE, SimWinchBrakeOpenDelayS := 0.042, RawPosM1 := RawPosM1, RawPosM2 := RawPosM2);
    ASSERT_TRUE(FB_Bench.Winch.M1_BrakeIsOpen_DI, 'Delai ecoule (5e scan) : M1_BrakeIsOpen_DI bascule TRUE');
END_TEST

TEST 'TC-T300-INT-010 SimBench M3 publie le retour dynamique du drive'
VAR
    i : INT;
END_VAR
    FB_Bench(Enable := TRUE, M3_ReqTremie := TRUE, M3_ReqMaintenance := FALSE,
             M3_SpeedCmd_Pct := 50.0, M3_BrakeCmd := TRUE,
             RawPosM1 := RawPosM1, RawPosM2 := RawPosM2);
    FOR i := 1 TO 20 DO
        FB_Bench(Enable := TRUE, M3_ReqTremie := TRUE, M3_ReqMaintenance := FALSE,
                 M3_SpeedCmd_Pct := 50.0, M3_BrakeCmd := TRUE,
                 RawPosM1 := RawPosM1, RawPosM2 := RawPosM2);
    END_FOR;
    ASSERT_EQ(FB_Bench.Translation.M3_StatusWord, 16#0087, 'M3 actif apres ouverture frein et retour frequence');
    FB_Bench(Enable := TRUE, M3_ReqTremie := FALSE, M3_ReqMaintenance := FALSE,
             M3_SpeedCmd_Pct := 0.0, M3_BrakeCmd := FALSE,
             RawPosM1 := RawPosM1, RawPosM2 := RawPosM2);
    FOR i := 1 TO 50 DO
        FB_Bench(Enable := TRUE, M3_ReqTremie := FALSE, M3_ReqMaintenance := FALSE,
                 M3_SpeedCmd_Pct := 0.0, M3_BrakeCmd := FALSE,
                 RawPosM1 := RawPosM1, RawPosM2 := RawPosM2);
    END_FOR;
    ASSERT_EQ(FB_Bench.Translation.M3_StatusWord, 16#0080, 'M3 arrete apres decroissance reelle de frequence');
END_TEST

TEST 'TC-T300-INT-030 Image SimBench relaye les DI M3 au decodeur production'
VAR
    Decoder : FB_Translation_PositionDecoder;
    HwInTranslation : ST_HwTranslation;
    i : INT;
END_VAR
    (* Le premier appel neutralise l'etat precedent. La copie explicite ci-dessous
       est representative du pont reel HwSim.Translation -> HwIn.Translation ;
       son unicite dans le programme est imposee statiquement par G502. *)
    FB_Bench(Enable := FALSE, RawPosM1 := RawPosM1, RawPosM2 := RawPosM2);
    FB_Bench(Enable := TRUE, M3_ReqTremie := FALSE, M3_ReqMaintenance := FALSE,
             M3_SpeedCmd_Pct := 0.0, M3_BrakeCmd := FALSE,
             RawPosM1 := RawPosM1, RawPosM2 := RawPosM2);
    HwInTranslation := FB_Bench.Translation;
    Decoder(SensorTremie := HwInTranslation.M3_PosTremie_DI,
            SensorPV := HwInTranslation.M3_PosPV_DI,
            SensorP2 := HwInTranslation.M3_PosPVP2_DI,
            SensorP1 := HwInTranslation.M3_PosP1_DI,
            SensorMaintenance := HwInTranslation.M3_PosMaintenance_DI);
    ASSERT_EQ(Decoder.SensorsWord, 2#00011, 'Repli P1 publie par l image puis decode sans injection aval');
    ASSERT_FALSE(Decoder.Incoherent, 'Mot P1 issu du SimBench coherent au decodeur production');

    (* T361 — 1800 scans (18 s) au lieu de 1100 : le banc a ete recale sur le gain odometrique
       reel (CST_M3FullTravelTimeS 8,0 -> 37,5 s, soit 0,8 m/s a 40 Hz au lieu de 3,75 m/s).
       Le trajet P1 (20 m) -> capteur Maintenance (29,95 m) demande desormais ~14 s
       (9,95 m a 0,8 m/s + ~2 s de rampe de frequence + ouverture du frein) : a 1100 scans le
       chariot n'atteignait plus la fin de course et le cas testait autre chose que son objet.
       Marge restante : ~4 s, soit ~3 m avant la butee mecanique. *)
    FOR i := 1 TO 1800 DO
        FB_Bench(Enable := TRUE, M3_ReqTremie := FALSE, M3_ReqMaintenance := TRUE,
                 M3_SpeedCmd_Pct := 100.0, M3_BrakeCmd := TRUE,
                 RawPosM1 := RawPosM1, RawPosM2 := RawPosM2);
        HwInTranslation := FB_Bench.Translation;
        Decoder(SensorTremie := HwInTranslation.M3_PosTremie_DI,
                SensorPV := HwInTranslation.M3_PosPV_DI,
                SensorP2 := HwInTranslation.M3_PosPVP2_DI,
                SensorP1 := HwInTranslation.M3_PosP1_DI,
                SensorMaintenance := HwInTranslation.M3_PosMaintenance_DI);
    END_FOR;
    ASSERT_EQ(Decoder.SensorsWord, 2#00000, 'Fin Maintenance dynamique traverse image et decodeur');
    ASSERT_TRUE(Decoder.LimitSwitchMaintenance, 'FDC Maintenance derive uniquement du mot image');
    ASSERT_FALSE(Decoder.Incoherent, 'Fin Maintenance dynamique reste coherente');
END_TEST

TEST 'TC-T300-INT-031 Intermittence P1 dynamique relayee au decodeur production'
VAR
    Decoder : FB_Translation_PositionDecoder;
    HwInTranslation : ST_HwTranslation;
    P1Previous : BOOL;
    P1Lost : BOOL := FALSE;
    P1Recovered : BOOL := FALSE;
    i : INT;
END_VAR
    FB_Bench(Enable := FALSE, RawPosM1 := RawPosM1, RawPosM2 := RawPosM2);
    FB_Bench(Enable := TRUE, M3_ReqTremie := FALSE, M3_ReqMaintenance := FALSE,
             M3_SpeedCmd_Pct := 0.0, M3_BrakeCmd := FALSE,
             RawPosM1 := RawPosM1, RawPosM2 := RawPosM2);
    HwInTranslation := FB_Bench.Translation;
    P1Previous := HwInTranslation.M3_PosP1_DI;

    (* Angle declencheur nul : l'episode est impose par la traversee mecanique,
       pas par un mot DI force. La graine et la periode restent deterministes. *)
    FOR i := 1 TO 1500 DO
        FB_Bench(Enable := TRUE, M3_ReqTremie := FALSE, M3_ReqMaintenance := TRUE,
                 M3_SpeedCmd_Pct := 100.0, M3_BrakeCmd := TRUE,
                 SimM3SensorIntermittenceActive := TRUE,
                 SimM3SensorStabilizationS := 1.0,
                 SimM3SensorIntermittencePeriodS := 0.12,
                 SimM3SensorElectricalDelayS := 0.0,
                 SimM3SensorLoadAngleTriggerRad := 0.0,
                 SimM3SensorScenarioSeed := 3001,
                 RawPosM1 := RawPosM1, RawPosM2 := RawPosM2);
        HwInTranslation := FB_Bench.Translation;
        Decoder(SensorTremie := HwInTranslation.M3_PosTremie_DI,
                SensorPV := HwInTranslation.M3_PosPV_DI,
                SensorP2 := HwInTranslation.M3_PosPVP2_DI,
                SensorP1 := HwInTranslation.M3_PosP1_DI,
                SensorMaintenance := HwInTranslation.M3_PosMaintenance_DI);
        IF P1Previous AND NOT HwInTranslation.M3_PosP1_DI THEN
            P1Lost := TRUE;
        END_IF;
        IF P1Lost AND HwInTranslation.M3_PosP1_DI THEN
            P1Recovered := TRUE;
        END_IF;
        P1Previous := HwInTranslation.M3_PosP1_DI;
    END_FOR;
    ASSERT_TRUE(P1Lost, 'P1 perd au moins une fois son etat pendant le franchissement');
    ASSERT_TRUE(P1Recovered, 'P1 est repris pendant l episode borne');
    ASSERT_FALSE(HwInTranslation.M3_PosP1_DI, 'P1 se stabilise a FALSE apres franchissement vers Maintenance');
    ASSERT_FALSE(Decoder.TranslationPosP1, 'Decodeur production voit la stabilisation du DI image');
END_TEST

TEST 'T196-003 Capteur haut manuel et polarite Free_DI correcte'
    FB_Bench(Enable := TRUE, SimTopPositionActive := TRUE,
             RawPosM1 := RawPosM1, RawPosM2 := RawPosM2);
    ASSERT_FALSE(FB_Bench.Winch.M1M2_TopPositionFree_DI,
                 'TopPositionActive=TRUE -> Free_DI=FALSE (capteur atteint)');
    ADVANCE_TIME(10000000);
    FB_Bench(Enable := TRUE, SimTopPositionActive := FALSE,
             RawPosM1 := RawPosM1, RawPosM2 := RawPosM2);
    ASSERT_TRUE(FB_Bench.Winch.M1M2_TopPositionFree_DI,
                'TopPositionActive=FALSE -> Free_DI=TRUE (butée libre)');
END_TEST

TEST 'T196-004 Capteur haut auto : forçage manuel SimTopPositionActive'
    FB_Bench(Enable := TRUE, SimTopPositionActive := FALSE,
             RawPosM1 := RawPosM1, RawPosM2 := RawPosM2);
    ASSERT_TRUE(FB_Bench.Winch.M1M2_TopPositionFree_DI,
                'SimTopPositionActive=FALSE -> capteur haut libre');
    ADVANCE_TIME(10000000);
    FB_Bench(Enable := TRUE, SimTopPositionActive := TRUE,
             RawPosM1 := RawPosM1, RawPosM2 := RawPosM2);
    ASSERT_FALSE(FB_Bench.Winch.M1M2_TopPositionFree_DI,
                 'SimTopPositionActive=TRUE -> capteur haut actif');
END_TEST

(* =========================================================================
   AF-13 — FB_Sim_Safety (TC-P13-020/021/022/023)
   ========================================================================= *)

TEST 'TC-P13-020 Sim_Safety SimChainOk = A AND B AND NOT BtnEmergencyStop'
    FB_SimSafe(Enable := TRUE, SimChainOkBit := TRUE, BtnEmergencyStop := FALSE);
    ADVANCE_TIME(60000000); (* Delai retombe relais 50ms *)
    FB_SimSafe(Enable := TRUE, SimChainOkBit := TRUE, BtnEmergencyStop := FALSE);
    ASSERT_TRUE(FB_SimSafe.SimChainOk, 'SimChainOkBit=TRUE -> SimChainOk=TRUE apres 50ms');

    ADVANCE_TIME(10000000);
    FB_SimSafe(Enable := TRUE, SimChainOkBit := FALSE, BtnEmergencyStop := FALSE);
    ADVANCE_TIME(60000000);
    FB_SimSafe(Enable := TRUE, SimChainOkBit := FALSE, BtnEmergencyStop := FALSE);
    ASSERT_FALSE(FB_SimSafe.SimChainOk, 'SimChainOkBit=FALSE -> SimChainOk=FALSE');

    ADVANCE_TIME(10000000);
    FB_SimSafe(Enable := TRUE, SimChainOkBit := TRUE, BtnEmergencyStop := TRUE);
    ADVANCE_TIME(60000000);
    FB_SimSafe(Enable := TRUE, SimChainOkBit := TRUE, BtnEmergencyStop := TRUE);
    ASSERT_FALSE(FB_SimSafe.SimChainOk, 'BtnEmergencyStop -> SimChainOk=FALSE');
END_TEST

TEST 'TC-P13-021 Sim_Safety SimContactorOk s auto-maintient sur EmergencyArming'
    FB_SimSafe(Enable := TRUE, SimChainOkBit := TRUE, EmergencyArming := FALSE, BtnEmergencyStop := FALSE);
    ADVANCE_TIME(60000000);
    FB_SimSafe(Enable := TRUE, SimChainOkBit := TRUE, EmergencyArming := FALSE, BtnEmergencyStop := FALSE);
    ASSERT_FALSE(FB_SimSafe.SimContactorOk, 'pas encore arme -> contacteur FALSE');

    (* Impulsion armement tenue 100ms *)
    ADVANCE_TIME(10000000);
    FB_SimSafe(Enable := TRUE, SimChainOkBit := TRUE, EmergencyArming := TRUE, BtnEmergencyStop := FALSE);
    ADVANCE_TIME(110000000);
    FB_SimSafe(Enable := TRUE, SimChainOkBit := TRUE, EmergencyArming := TRUE, BtnEmergencyStop := FALSE);
    ASSERT_TRUE(FB_SimSafe.SimContactorOk, 'EmergencyArming -> contacteur engage');

    (* Relachement impulsion -> auto-maintien *)
    ADVANCE_TIME(10000000);
    FB_SimSafe(Enable := TRUE, SimChainOkBit := TRUE, EmergencyArming := FALSE, BtnEmergencyStop := FALSE);
    ASSERT_TRUE(FB_SimSafe.SimContactorOk, 'auto-maintien : contacteur reste engage');

    (* Coupure chaine -> retombe apres chaine (50ms) + contacteur (50ms) *)
    ADVANCE_TIME(10000000);
    FB_SimSafe(Enable := TRUE, SimChainOkBit := FALSE, EmergencyArming := FALSE, BtnEmergencyStop := FALSE);
    ADVANCE_TIME(60000000); (* Chaine s ouvre *)
    FB_SimSafe(Enable := TRUE, SimChainOkBit := FALSE, EmergencyArming := FALSE, BtnEmergencyStop := FALSE);
    ADVANCE_TIME(60000000); (* Contacteur retombe *)
    FB_SimSafe(Enable := TRUE, SimChainOkBit := FALSE, EmergencyArming := FALSE, BtnEmergencyStop := FALSE);
    ASSERT_FALSE(FB_SimSafe.SimContactorOk, 'SimChainOk=FALSE -> contacteur retombe');
END_TEST

TEST 'TC-P13-022 Sim_Safety Enable=FALSE neutralise tout'
    FB_SimSafe(Enable := FALSE, PowerCutOff_A := TRUE, PowerCutOff_B := TRUE, EmergencyArming := TRUE, BtnEmergencyStop := FALSE);
    ASSERT_FALSE(FB_SimSafe.SimChainOk, 'Enable=FALSE -> SimChainOk=FALSE');
    ASSERT_FALSE(FB_SimSafe.SimContactorOk, 'Enable=FALSE -> SimContactorOk=FALSE');
END_TEST

TEST 'TC-P13-023 Sim_Safety latch AU non lie a la sim (essai manuel — stub)'
    (* Stub : TC-P13-023 verifie qu un defaut AU reel latche (RedundancyTestFailedCause /
       EmergencyArmingFailedCause dans FB_Safety_EmergencyManagementLogic) survit a la sim et
       ne se debloque que par front Reset runtime. Non automatisable en boite noire FB_Sim_Safety
       (latch dans le FB consommateur). (essai manuel — stub) *)
    ASSERT_TRUE(TRUE, 'Stub : latch AU a verifier manuellement (essai manuel)');
END_TEST

(* =========================================================================
   AF-13 — FB_Sim_Encoder (TC-P13-030/031/032/033)
   ========================================================================= *)

TEST 'TC-P13-030 Sim_Encoder RelayFwd/Rev font compter RawPos'
    RawPosM1 := 0;
    FB_SimEnc(Enable := TRUE, RelayFwd := TRUE, RelayRev := FALSE, StepNumber := 1, RawPos := RawPosM1);
    ASSERT_GT(FB_SimEnc.RawPosOut, 0, 'RelayFwd -> RawPos augmente');
    ADVANCE_TIME(10000000);
    RawPosM1 := 100;
    FB_SimEnc(Enable := TRUE, RelayFwd := TRUE, RelayRev := FALSE, StepNumber := 1, RawPos := RawPosM1);
    ASSERT_GT(FB_SimEnc.RawPosOut, 100, 'RelayFwd -> RawPos augmente depuis 100');
    ADVANCE_TIME(10000000);
    RawPosM1 := 100;
    FB_SimEnc(Enable := TRUE, RelayFwd := FALSE, RelayRev := TRUE, StepNumber := 1, RawPos := RawPosM1);
    ASSERT_LT(FB_SimEnc.RawPosOut, 100, 'RelayRev -> RawPos diminue');
END_TEST

TEST 'TC-P13-031 Sim_Encoder PresetCmd charge PresetValue'
    RawPosM1 := 0;
    FB_SimEnc(Enable := TRUE, RelayFwd := FALSE, RelayRev := FALSE, StepNumber := 1, PresetCmd := TRUE, PresetValue := 5000, RawPos := RawPosM1);
    ADVANCE_TIME(10000000);
    FB_SimEnc(Enable := TRUE, RelayFwd := FALSE, RelayRev := FALSE, StepNumber := 1, PresetCmd := FALSE, PresetValue := 5000, RawPos := RawPosM1);
    ADVANCE_TIME(10000000);
    FB_SimEnc(Enable := TRUE, RelayFwd := FALSE, RelayRev := FALSE, StepNumber := 1, PresetCmd := FALSE, PresetValue := 5000, RawPos := RawPosM1);
    ADVANCE_TIME(10000000);
    FB_SimEnc(Enable := TRUE, RelayFwd := FALSE, RelayRev := FALSE, StepNumber := 1, PresetCmd := FALSE, PresetValue := 5000, RawPos := RawPosM1);
    ASSERT_EQ(FB_SimEnc.RawPosOut, 5000, 'Preset applique apres latence');
END_TEST

TEST 'TC-P13-032 Sim_Encoder le comptage franchit 0 au lieu de s y figer (butee silencieuse supprimee, T338)'
    (* Realigne sur la semantique T338 (comptage brut SIGNED 32 bits) : cette copie etait restee
       sur l'ancienne butee `RawPos := 0`, ce qui rendait la suite FB_SimBench ROUGE (41/42) sur
       HEAD depuis le commit 6a5910da — non-regression T338 incomplete. *)
    RawPosM1 := 41; (* 41 pts = exactement un pas de descente au palier 1 (1,0 x 4096 x 0,010) *)
    FB_SimEnc(Enable := TRUE, RelayFwd := FALSE, RelayRev := TRUE, StepNumber := 1, RawPos := RawPosM1);
    RawPosM1 := FB_SimEnc.RawPosOut; (* le caller conserve la memoire persistante du codeur *)
    ASSERT_EQ(FB_SimEnc.RawPosOut, 0, 'Un pas de descente amene le comptage exactement a 0 (point de passage)');
    ADVANCE_TIME(10000000);
    FB_SimEnc(Enable := TRUE, RelayFwd := FALSE, RelayRev := TRUE, StepNumber := 1, RawPos := RawPosM1);
    RawPosM1 := FB_SimEnc.RawPosOut;
    ASSERT_TRUE(FB_SimEnc.RawPosOut <> 0, 'Scan suivant : le comptage franchit 0 au lieu de s y figer');
    ASSERT_EQ(FB_SimEnc.RawPosOut, 4294967255, 'Comptage = -41 pts (aucune borne a 0, 2^32 - 41 en signe)');
END_TEST

TEST 'TC-P13-033 Sim_Encoder RawPos survit a un reset froid (essai manuel — stub)'
    (* Stub : TC-P13-033 verifie que RawPos (VAR_IN_OUT reference GVL_PERSISTENT) survit a un
       reset froid. Non automatisable en boite noire (depend de la persistance CODESYS).
       (essai manuel — stub) *)
    ASSERT_TRUE(TRUE, 'Stub : persistance RawPos a verifier manuellement (essai manuel)');
END_TEST

(* =========================================================================
   AF-13 — FB_Sim_Translation (TC-P13-040/041/042/043)
   ========================================================================= *)

TEST 'TC-T300-INT-020 Sim_Translation initialise le mot P1'
    FB_SimTrans(Enable := TRUE, ReqTremie := FALSE, ReqMaintenance := FALSE,
                SpeedTgt_Pct := 0.0, BrakeReleaseCmd := FALSE);
    ASSERT_FALSE(FB_SimTrans.PosTremie, 'P1 ne doit pas annoncer Tremie');
    ASSERT_FALSE(FB_SimTrans.PosPV, 'P1 ne doit pas annoncer PV');
    ASSERT_FALSE(FB_SimTrans.PosP2, 'P1 ne doit pas annoncer P2');
    ASSERT_TRUE(FB_SimTrans.PosP1, 'P1 actif au repli');
    ASSERT_TRUE(FB_SimTrans.PosMaintenance, 'Mot thermometre P1 coherent');
END_TEST

TEST 'TC-T300-INT-021 Sim_Translation neutralise deux sens simultanes'
    FB_SimTrans(Enable := TRUE, ReqTremie := TRUE, ReqMaintenance := TRUE,
                SpeedTgt_Pct := 100.0, BrakeReleaseCmd := TRUE);
    ASSERT_EQ(FB_SimTrans.FrequencyCmd_Hz, 0.0, 'Deux sens ne creent aucune consigne');
    ASSERT_EQ(FB_SimTrans.ActualFrequency_Hz, 0.0, 'Aucun retour variateur sans sens unique');
END_TEST

TEST 'TC-T300-INT-022 Sim_Translation borne et publie la fin de course Maintenance'
VAR
    i : INT;
END_VAR
    FB_SimTrans(Enable := FALSE);
    FB_SimTrans(Enable := TRUE, ReqTremie := FALSE, ReqMaintenance := TRUE,
                SpeedTgt_Pct := 100.0, FullTravelTimeS := 0.5,
                BrakeReleaseCmd := TRUE, SensorElectricalDelayS := 0.0);
    FOR i := 1 TO 400 DO
        FB_SimTrans(Enable := TRUE, ReqTremie := FALSE, ReqMaintenance := TRUE,
                    SpeedTgt_Pct := 100.0, FullTravelTimeS := 0.5,
                    BrakeReleaseCmd := TRUE, SensorElectricalDelayS := 0.0);
    END_FOR;
    ASSERT_GE(FB_SimTrans.PositionTrue_M, 0.0, 'Borne Tremie respectee');
    ASSERT_LE(FB_SimTrans.PositionTrue_M, 30.0, 'Borne Maintenance respectee');
    ASSERT_FALSE(FB_SimTrans.PosMaintenance, 'Maintenance publie le mot 00000 a la butee');
END_TEST

TEST 'TC-T300-INT-023 Sim_Translation desactive se replie P1'
    FB_SimTrans(Enable := FALSE, ReqTremie := FALSE, ReqMaintenance := TRUE,
                SpeedTgt_Pct := 100.0, BrakeReleaseCmd := TRUE);
    ASSERT_EQ(FB_SimTrans.PositionTrue_M, 20.0, 'Repli physique P1');
    ASSERT_TRUE(FB_SimTrans.PosP1, 'Capteur P1 coherent hors simulation');
    ASSERT_TRUE(FB_SimTrans.PosMaintenance, 'Mot P1 coherent hors simulation');
    ASSERT_FALSE(FB_SimTrans.BrakeContactOpen, 'Frein confirme ferme hors simulation');
END_TEST

(* =========================================================================
   AF-13 — FB_Sim_Joystick (TC-P13-050/051/052)
   ========================================================================= *)

TEST 'TC-P13-050 Sim_Joystick initialise au neutre au premier cycle'
    FB_SimJoy(Enable := TRUE, NeutralRaw := 5000, MaxRaw := 10000);
    ASSERT_EQ(FB_SimJoy.RawX, 5000, 'premier cycle -> RawX=NeutralRaw');
    ASSERT_EQ(FB_SimJoy.RawY, 5000, 'premier cycle -> RawY=NeutralRaw');
    ASSERT_FALSE(FB_SimJoy.RawButton, 'premier cycle -> RawButton=FALSE');
END_TEST

TEST 'TC-P13-051 Sim_Joystick sorties forçables en instance (essai manuel — stub)'
    (* Stub : TC-P13-051 verifie que RawX/RawY/RawButton restent forçables librement en instance
       CODESYS apres l'init (le FB n'ecrit plus ces sorties apres le premier cycle). Non
       automatisable en boite noire (depend du forçage CODESYS). (essai manuel — stub) *)
    ASSERT_TRUE(TRUE, 'Stub : forçage joystick a verifier manuellement (essai manuel)');
END_TEST

TEST 'TC-P13-052 Sim_Joystick homme-mort : RawButton reflete l appui (partie AUTO)'
    (* Aucun bouton -> RawButton=FALSE *)
    FB_SimJoy(Enable := TRUE, NeutralRaw := 5000, MaxRaw := 10000);
    ASSERT_FALSE(FB_SimJoy.RawButton, 'aucun bouton -> RawButton=FALSE');
    ADVANCE_TIME(10000000);
    (* Bouton directionnel actif -> RawButton=TRUE (homme-mort inclus) *)
    FB_SimJoy(Enable := TRUE, NeutralRaw := 5000, MaxRaw := 10000, BtnRight_Fwd_MAINT := TRUE);
    ASSERT_TRUE(FB_SimJoy.RawButton, 'bouton actif -> RawButton=TRUE');
END_TEST

(* =========================================================================
   AF-13 — FB_SimBench : rattrapage mecanique M1/M2 (T328)
   Plan : DOC/WFLOW/CONTRACTS/PLAN_T328_SIMBENCH_COUPLAGE_MECANIQUE_M1M2.md
   ========================================================================= *)

TEST 'TC-P13-060 T328 montee couplee : rattrapage actif et correction bornee'
    (* Montée couplée réelle (relais M1+M2 même sens, freins desserrés), benne DANS le trou métier
       T327 : écart 13,5 m < entrée de bande fermée (14,5 m). Le rattrapage agit, borné par la pente. *)
    RawPosM1 := 1000000; RawPosM2 := 1100000;
    FB_Bench(Enable := TRUE, RawPosM1 := RawPosM1, RawPosM2 := RawPosM2,
             M1_RelayFwd := TRUE, M2_RelayFwd := TRUE,
             M1_BrakeCmd := TRUE, M2_BrakeCmd := TRUE,
             SimWinchCouplingModelActive := TRUE,
             M1_CablePos_M := 5.0, M2_CablePos_M := 18.5,
             BucketOffsetCloseM := 15.0, BucketCoherenceLimitM := 1.0);
    ASSERT_TRUE(FB_Bench.WinchCouplingActive, 'montee couplee -> rattrapage actif');
    ASSERT_TRUE(FB_Bench.WinchCouplingCorrectionPts > 0, 'ecart sous la bande -> correction non nulle');
    ASSERT_TRUE(FB_Bench.WinchCouplingCorrectionPts <= 82, 'correction bornee (0,02 m/scan = 82 points)');
    ASSERT_TRUE(FB_Bench.Winch.COD2_PosValue > RawPosM2, 'correction appliquee a l IMAGE M2 uniquement');
END_TEST

TEST 'TC-P13-061 T328 arret et jog M2 seul : ecart fige, aucune correction'
    (* Relais à 0 : aucun mouvement réel -> jamais de rattrapage (AC6). *)
    FB_Bench(Enable := TRUE, RawPosM1 := RawPosM1, RawPosM2 := RawPosM2,
             M1_RelayFwd := FALSE, M2_RelayFwd := FALSE,
             SimWinchCouplingModelActive := TRUE,
             M1_CablePos_M := 5.0, M2_CablePos_M := 18.5,
             BucketOffsetCloseM := 15.0, BucketCoherenceLimitM := 1.0);
    ASSERT_FALSE(FB_Bench.WinchCouplingActive, 'relais a 0 -> pas de rattrapage');
    ASSERT_EQ(FB_Bench.WinchCouplingCorrectionPts, 0, 'aucune correction a l arret');
    ASSERT_EQ(FB_Bench.Winch.COD2_PosValue, RawPosM2, 'image M2 inchangee a l arret');
    ADVANCE_TIME(10000000);
    (* Jog M2 seul (un seul treuil actif) -> toujours aucun rattrapage *)
    FB_Bench(Enable := TRUE, RawPosM1 := RawPosM1, RawPosM2 := RawPosM2,
             M1_RelayFwd := FALSE, M2_RelayFwd := TRUE,
             M1_BrakeCmd := FALSE, M2_BrakeCmd := TRUE,
             SimWinchCouplingModelActive := TRUE,
             M1_CablePos_M := 5.0, M2_CablePos_M := 18.5,
             BucketOffsetCloseM := 15.0, BucketCoherenceLimitM := 1.0);
    ASSERT_FALSE(FB_Bench.WinchCouplingActive, 'jog M2 seul -> pas de rattrapage');
    ASSERT_EQ(FB_Bench.WinchCouplingCorrectionPts, 0, 'jog M2 seul -> aucune correction');
END_TEST

TEST 'TC-P13-062 T328 machoires bloquees : rattrapage inhibe et charge forcee'
    FB_Bench(Enable := TRUE, RawPosM1 := RawPosM1, RawPosM2 := RawPosM2,
             M1_RelayFwd := TRUE, M2_RelayFwd := TRUE,
             M1_BrakeCmd := TRUE, M2_BrakeCmd := TRUE,
             SimWinchCouplingModelActive := TRUE,
             SimBucketJamActive := TRUE,
             SimWinchElectricalDiagnosticsActive := TRUE,
             M1_CablePos_M := 5.0, M2_CablePos_M := 18.5,
             BucketOffsetCloseM := 15.0, BucketCoherenceLimitM := 1.0);
    ASSERT_FALSE(FB_Bench.WinchCouplingActive, 'blocage machoires -> rattrapage inhibe');
    ASSERT_EQ(FB_Bench.WinchCouplingCorrectionPts, 0, 'blocage -> aucune correction');
    ASSERT_TRUE(FB_Bench.MotorTorqueM1_Nm > 0.0, 'blocage -> charge forcee observable (diagnostic)');
END_TEST

TEST 'TC-P13-063 T328 modele desactive : image M2 inchangee (non-masquage T327)'
    FB_Bench(Enable := TRUE, RawPosM1 := RawPosM1, RawPosM2 := RawPosM2,
             M1_RelayFwd := TRUE, M2_RelayFwd := TRUE,
             M1_BrakeCmd := TRUE, M2_BrakeCmd := TRUE,
             SimWinchCouplingModelActive := FALSE,
             M1_CablePos_M := 5.0, M2_CablePos_M := 18.5,
             BucketOffsetCloseM := 15.0, BucketCoherenceLimitM := 1.0);
    ASSERT_FALSE(FB_Bench.WinchCouplingActive, 'modele OFF -> pas de rattrapage');
    ASSERT_EQ(FB_Bench.WinchCouplingCorrectionPts, 0, 'modele OFF -> aucune correction');
    ASSERT_EQ(FB_Bench.Winch.COD2_PosValue, RawPosM2, 'modele OFF -> image M2 identique (trou T327 preserve)');
END_TEST

TEST 'TC-P13-064 T328 cable mou : rattrapage inhibe (aucun effort transmis)'
    FB_Bench(Enable := TRUE, RawPosM1 := RawPosM1, RawPosM2 := RawPosM2,
             M1_RelayFwd := TRUE, M2_RelayFwd := TRUE,
             M1_BrakeCmd := TRUE, M2_BrakeCmd := TRUE,
             SimWinchCouplingModelActive := TRUE,
             SimM2TensionedCableFaultInject := TRUE,
             M1_CablePos_M := 5.0, M2_CablePos_M := 18.5,
             BucketOffsetCloseM := 15.0, BucketCoherenceLimitM := 1.0);
    ASSERT_FALSE(FB_Bench.WinchCouplingActive, 'cable mou -> pas de rattrapage');
END_TEST

TEST 'TC-P13-065 T328 banc eteint : image reelle repliquee sans correction'
    FB_Bench(Enable := FALSE, RawPosM1 := RawPosM1, RawPosM2 := RawPosM2,
             M1_RelayFwd := TRUE, M2_RelayFwd := TRUE,
             M1_BrakeCmd := TRUE, M2_BrakeCmd := TRUE,
             SimWinchCouplingModelActive := TRUE,
             M1_CablePos_M := 5.0, M2_CablePos_M := 18.5,
             BucketOffsetCloseM := 15.0, BucketCoherenceLimitM := 1.0);
    ASSERT_FALSE(FB_Bench.WinchCouplingActive, 'banc desactive -> aucun rattrapage');
    ASSERT_EQ(FB_Bench.Winch.COD2_PosValue, RawPosM2, 'banc desactive -> image sans correction');
END_TEST

TEST 'TC-P13-066 T328 convergence multi-scan du rattrapage vers la bande fermee'
VAR
    i        : INT;
    M2_Pos_M : REAL := 0.0;
END_VAR
    (* Boucle fermee simulee : la position M2 vue par le metier suit l'image corrigee, comme dans la
       chaine reelle (HwSim -> HwIn -> codeur). Delta initial 13,5 m = trou metier de fermeture.
       Chaque appel du FB vaut un scan de 10 ms (le modele utilise CST_SimBenchCycleTimeS, pas le
       temps du harness) : la boucle n'avance donc pas le temps du harness. *)
    RawPosM1 := 1000000; RawPosM2 := 1100000;
    M2_Pos_M := 18.5;   (* Delta = M2 - M1 = 13,5 m *)
    FOR i := 1 TO 100 DO
        FB_Bench(Enable := TRUE, RawPosM1 := RawPosM1, RawPosM2 := RawPosM2,
                 M1_RelayFwd := TRUE, M2_RelayFwd := TRUE,
                 M1_BrakeCmd := TRUE, M2_BrakeCmd := TRUE,
                 SimWinchCouplingModelActive := TRUE,
                 M1_CablePos_M := 5.0, M2_CablePos_M := M2_Pos_M,
                 BucketOffsetCloseM := 15.0, BucketCoherenceLimitM := 1.0);
        ASSERT_TRUE(FB_Bench.WinchCouplingCorrectionPts <= 82, 'correction bornee a 0,02 m par scan');
        M2_Pos_M := M2_Pos_M + DINT_TO_REAL(FB_Bench.WinchCouplingCorrectionPts) * (2.0 / 8192.0);
    END_FOR;
    ADVANCE_TIME(10000000);
    ASSERT_TRUE((M2_Pos_M - 5.0) >= 14.0, 'Delta entre dans la bande fermee (>= 14,0 m) en temps borne');
END_TEST

TEST 'TC-P13-067 T328 un preset purge l offset de reprise de jeu (image = codeur)'
    RawPosM1 := 1000000; RawPosM2 := 1100000;
    (* Session active : un offset est bien accumule. *)
    FB_Bench(Enable := TRUE, RawPosM1 := RawPosM1, RawPosM2 := RawPosM2,
             M1_RelayFwd := TRUE, M2_RelayFwd := TRUE,
             M1_BrakeCmd := TRUE, M2_BrakeCmd := TRUE,
             SimWinchCouplingModelActive := TRUE,
             M1_CablePos_M := 5.0, M2_CablePos_M := 18.5,
             BucketOffsetCloseM := 15.0, BucketCoherenceLimitM := 1.0);
    ASSERT_TRUE(FB_Bench.Winch.COD2_PosValue > RawPosM2, 'offset de reprise de jeu accumule');
    ADVANCE_TIME(10000000);
    (* Preset M2 (PresetTriggerCmd = 2) : la reference absolue est reecrite -> offset purge. *)
    FB_Bench(Enable := TRUE, RawPosM1 := RawPosM1, RawPosM2 := RawPosM2,
             M1_RelayFwd := TRUE, M2_RelayFwd := TRUE,
             M1_BrakeCmd := TRUE, M2_BrakeCmd := TRUE,
             SimWinchCouplingModelActive := TRUE, M2_PresetTriggerCmd := 2,
             M1_CablePos_M := 5.0, M2_CablePos_M := 18.5,
             BucketOffsetCloseM := 15.0, BucketCoherenceLimitM := 1.0);
    ASSERT_EQ(FB_Bench.Winch.COD2_PosValue, RawPosM2, 'preset -> offset purge, image = codeur');
END_TEST

TEST 'TC-P13-068 T328 mode OFF apres session active : aucun offset residuel'
    RawPosM1 := 1000000; RawPosM2 := 1100000;
    FB_Bench(Enable := TRUE, RawPosM1 := RawPosM1, RawPosM2 := RawPosM2,
             M1_RelayFwd := TRUE, M2_RelayFwd := TRUE,
             M1_BrakeCmd := TRUE, M2_BrakeCmd := TRUE,
             SimWinchCouplingModelActive := TRUE,
             M1_CablePos_M := 5.0, M2_CablePos_M := 18.5,
             BucketOffsetCloseM := 15.0, BucketCoherenceLimitM := 1.0);
    ASSERT_TRUE(FB_Bench.Winch.COD2_PosValue > RawPosM2, 'offset accumule en mode actif');
    ADVANCE_TIME(10000000);
    (* Bascule mode OFF : l'image doit redevenir strictement celle du codeur (non-masquage). *)
    FB_Bench(Enable := TRUE, RawPosM1 := RawPosM1, RawPosM2 := RawPosM2,
             M1_RelayFwd := TRUE, M2_RelayFwd := TRUE,
             M1_BrakeCmd := TRUE, M2_BrakeCmd := TRUE,
             SimWinchCouplingModelActive := FALSE,
             M1_CablePos_M := 5.0, M2_CablePos_M := 18.5,
             BucketOffsetCloseM := 15.0, BucketCoherenceLimitM := 1.0);
    ASSERT_FALSE(FB_Bench.WinchCouplingActive, 'mode OFF -> rattrapage inactif');
    ASSERT_EQ(FB_Bench.Winch.COD2_PosValue, RawPosM2, 'mode OFF -> aucun offset residuel sur l image');
END_TEST

(* =========================================================================
   T328 (reprise DSH03) — SCENARIO UTILISATEUR 2026-09-20 : benne FERMEE avec
   ecart residuel ~5 % (voyant ferme allume), puis MONTEE couplee.
   Definitions (source FB_Bucket.st:591 + GVL_PERSISTENT.st:66-70) :
     Ouverture_Pct = 100 * (OffsetCloseM - Delta) / (OffsetCloseM - OffsetOpenM)
     Delta = CablePosM2 - CablePosM1 ; OffsetCloseM = 15,0 m ; OffsetOpenM = 0,0 m
     => ecart 5 %  <=> Delta = 14,25 m   (=> IsClosed TRUE : Delta >= 14,0 m)
        ecart 0 %  <=> Delta = 15,0 m   (butee mecanique benne fermee)
        ecart 3,33 % <=> Delta = 14,50 m (cible ABANDONNEE (plafonnait l ecart a 3,4 %), FB_SimBench.st:505)
   Aucun de ces cas n existait dans la suite : TC-P13-060..068 partent tous de
   Delta = 13,5 m (10 % ouverture, trou metier T327), jamais du residuel POST-fermeture.
   CIBLE RETENUE (arbitrage CC01 2026-09-20, D1) : BUTEE mecanique (ecart 0 %).
   ========================================================================= *)

TEST 'TC-P13-070 T328 scenario utilisateur : ecart 5 % (Delta 14,25 m) resorbe vers 0 % en montee couplee'
VAR
    i        : INT;
    M2_Pos_M : REAL := 0.0;
END_VAR
    (* Boucle fermee reelle : HwSim (image corrigee) -> HwIn -> codeur M2 -> Delta mesure. *)
    RawPosM1 := 1000000; RawPosM2 := 1100000;
    M2_Pos_M := 14.25 + 5.0;   (* Delta initial = 14,25 m => ouverture 5 % (cas utilisateur) *)
    FOR i := 1 TO 800 DO
        FB_Bench(Enable := TRUE, RawPosM1 := RawPosM1, RawPosM2 := RawPosM2,
                 M1_RelayFwd := TRUE, M2_RelayFwd := TRUE,
                 M1_BrakeCmd := TRUE, M2_BrakeCmd := TRUE,
                 SimWinchCouplingModelActive := TRUE,
                 M1_CablePos_M := 5.0, M2_CablePos_M := M2_Pos_M,
                 BucketOffsetCloseM := 15.0, BucketCoherenceLimitM := 1.0);
        ASSERT_TRUE(FB_Bench.WinchCouplingCorrectionPts <= 82, 'correction bornee a 0,02 m par scan');
        M2_Pos_M := M2_Pos_M + DINT_TO_REAL(FB_Bench.WinchCouplingCorrectionPts) * (2.0 / 8192.0);
    END_FOR;
    ADVANCE_TIME(10000000);
    (* Plancher de quantification : arret des que l increment < 1 point codeur (0,244 mm)
       => ecart residuel <= 2,5 cm soit 0,17 %, affiche 0 % a l IHM. *)
    ASSERT_TRUE((M2_Pos_M - 5.0) >= 14.97, 'ECART ATTENDU 0 % (Delta -> butee 15,0 m) pendant la montee');
    ASSERT_TRUE((M2_Pos_M - 5.0) <= 15.0, 'jamais de depassement de la butee mecanique');
END_TEST

TEST 'TC-P13-071 T328 cible : le point fixe du modele EST la butee mecanique (ecart 0 %)'
VAR
    i        : INT;
    M2_Pos_M : REAL := 0.0;
END_VAR
    (* Meme scenario que TC-P13-070 : on MESURE le point fixe du modele apres correctif D1.
       Cible = OffsetCloseM = 15,00 m ; point fixe mesure >= 14,975 m : le modele s arrete des que
       l increment 1er ordre devient < 1 point codeur (0,244 mm), soit un residu <= 2,5 cm.
       => ouverture residuelle <= 0,17 %, jamais un plancher de 3,4 %. *)
    RawPosM1 := 1000000; RawPosM2 := 1100000;
    M2_Pos_M := 14.25 + 5.0;
    FOR i := 1 TO 800 DO
        FB_Bench(Enable := TRUE, RawPosM1 := RawPosM1, RawPosM2 := RawPosM2,
                 M1_RelayFwd := TRUE, M2_RelayFwd := TRUE,
                 M1_BrakeCmd := TRUE, M2_BrakeCmd := TRUE,
                 SimWinchCouplingModelActive := TRUE,
                 M1_CablePos_M := 5.0, M2_CablePos_M := M2_Pos_M,
                 BucketOffsetCloseM := 15.0, BucketCoherenceLimitM := 1.0);
        M2_Pos_M := M2_Pos_M + DINT_TO_REAL(FB_Bench.WinchCouplingCorrectionPts) * (2.0 / 8192.0);
    END_FOR;
    ADVANCE_TIME(10000000);
    ASSERT_NEAR(M2_Pos_M - 5.0, 15.0, 0.03);
    ASSERT_TRUE((M2_Pos_M - 5.0) <= 15.0, 'point fixe = butee, jamais au-dela');
END_TEST

TEST 'TC-P13-072 T328 sur-fermeture (Delta > butee) : ecart FIGE, jamais corrige'
VAR
    i        : INT;
    M2_Pos_M : REAL := 0.0;
END_VAR
    (* Decision CC01 2026-09-20 (D2) : une sur-fermeture (Delta 15,75 m, soit +5 % AU-DELA de la
       butee 15,0 m, toujours dans la bande fermee 14,0..16,0 m) n est PAS corrigee : le modele
       reste strictement unidirectionnel -> rouvrir la benne pour resorber une sur-fermeture
       serait un mouvement non commande. Ecart FIGE : comportement voulu et teste. *)
    RawPosM1 := 1000000; RawPosM2 := 1100000;
    M2_Pos_M := 15.75 + 5.0;
    FOR i := 1 TO 100 DO
        FB_Bench(Enable := TRUE, RawPosM1 := RawPosM1, RawPosM2 := RawPosM2,
                 M1_RelayFwd := TRUE, M2_RelayFwd := TRUE,
                 M1_BrakeCmd := TRUE, M2_BrakeCmd := TRUE,
                 SimWinchCouplingModelActive := TRUE,
                 M1_CablePos_M := 5.0, M2_CablePos_M := M2_Pos_M,
                 BucketOffsetCloseM := 15.0, BucketCoherenceLimitM := 1.0);
        ASSERT_EQ(FB_Bench.WinchCouplingCorrectionPts, 0, 'sur-fermeture 5 % -> aucune correction');
        M2_Pos_M := M2_Pos_M + DINT_TO_REAL(FB_Bench.WinchCouplingCorrectionPts) * (2.0 / 8192.0);
    END_FOR;
    ADVANCE_TIME(10000000);
    ASSERT_NEAR(M2_Pos_M - 5.0, 15.75, 0.01);
END_TEST

TEST 'TC-P13-073 T328 GARDE-FOU : toute la bande de residus post-fermeture converge vers la butee'
VAR
    i        : INT;
    M2_Pos_M : REAL := 0.0;
END_VAR
    (* Garde-fou du trou de test qui a laisse passer T328 : la suite livree ne testait QUE
       Delta = 13,5 m. On couvre la bande des residus POST-fermeture reellement produite par la
       coupure d'anticipation + le roulis : 13,8 m (coupure T327) / 14,25 m (cas utilisateur 5 %) /
       14,75 m (haut de bande). Les trois doivent rejoindre la butee (ecart 0 %).
       (3 scenarios deroules : le harnais n accepte pas les boucles FOR imbriquees.) *)
    RawPosM1 := 1000000; RawPosM2 := 1100000;

    (* --- Residu 13,8 m (coupure d'anticipation T327) --- *)
    M2_Pos_M := 13.8 + 5.0;
    FOR i := 1 TO 800 DO
        FB_Bench(Enable := TRUE, RawPosM1 := RawPosM1, RawPosM2 := RawPosM2,
                 M1_RelayFwd := TRUE, M2_RelayFwd := TRUE,
                 M1_BrakeCmd := TRUE, M2_BrakeCmd := TRUE,
                 SimWinchCouplingModelActive := TRUE,
                 M1_CablePos_M := 5.0, M2_CablePos_M := M2_Pos_M,
                 BucketOffsetCloseM := 15.0, BucketCoherenceLimitM := 1.0);
        ASSERT_TRUE(FB_Bench.WinchCouplingCorrectionPts <= 82, 'correction bornee a 0,02 m par scan');
        M2_Pos_M := M2_Pos_M + DINT_TO_REAL(FB_Bench.WinchCouplingCorrectionPts) * (2.0 / 8192.0);
    END_FOR;
    ADVANCE_TIME(10000000);
    ASSERT_TRUE((M2_Pos_M - 5.0) >= 14.97, 'residu 13,8 m -> butee atteinte (ecart <= 0,2 %)');
    ASSERT_TRUE((M2_Pos_M - 5.0) <= 15.0, 'residu 13,8 m -> aucun depassement de butee');

    (* --- Residu 14,25 m (cas utilisateur : ecart 5 %, voyant ferme allume) --- *)
    M2_Pos_M := 14.25 + 5.0;
    FOR i := 1 TO 800 DO
        FB_Bench(Enable := TRUE, RawPosM1 := RawPosM1, RawPosM2 := RawPosM2,
                 M1_RelayFwd := TRUE, M2_RelayFwd := TRUE,
                 M1_BrakeCmd := TRUE, M2_BrakeCmd := TRUE,
                 SimWinchCouplingModelActive := TRUE,
                 M1_CablePos_M := 5.0, M2_CablePos_M := M2_Pos_M,
                 BucketOffsetCloseM := 15.0, BucketCoherenceLimitM := 1.0);
        ASSERT_TRUE(FB_Bench.WinchCouplingCorrectionPts <= 82, 'correction bornee a 0,02 m par scan');
        M2_Pos_M := M2_Pos_M + DINT_TO_REAL(FB_Bench.WinchCouplingCorrectionPts) * (2.0 / 8192.0);
    END_FOR;
    ADVANCE_TIME(10000000);
    ASSERT_TRUE((M2_Pos_M - 5.0) >= 14.97, 'residu 14,25 m -> butee atteinte (ecart <= 0,2 %)');
    ASSERT_TRUE((M2_Pos_M - 5.0) <= 15.0, 'residu 14,25 m -> aucun depassement de butee');

    (* --- Residu 14,75 m (haut de bande fermee) --- *)
    M2_Pos_M := 14.75 + 5.0;
    FOR i := 1 TO 800 DO
        FB_Bench(Enable := TRUE, RawPosM1 := RawPosM1, RawPosM2 := RawPosM2,
                 M1_RelayFwd := TRUE, M2_RelayFwd := TRUE,
                 M1_BrakeCmd := TRUE, M2_BrakeCmd := TRUE,
                 SimWinchCouplingModelActive := TRUE,
                 M1_CablePos_M := 5.0, M2_CablePos_M := M2_Pos_M,
                 BucketOffsetCloseM := 15.0, BucketCoherenceLimitM := 1.0);
        ASSERT_TRUE(FB_Bench.WinchCouplingCorrectionPts <= 82, 'correction bornee a 0,02 m par scan');
        M2_Pos_M := M2_Pos_M + DINT_TO_REAL(FB_Bench.WinchCouplingCorrectionPts) * (2.0 / 8192.0);
    END_FOR;
    ADVANCE_TIME(10000000);
    ASSERT_TRUE((M2_Pos_M - 5.0) >= 14.97, 'residu 14,75 m -> butee atteinte (ecart <= 0,2 %)');
    ASSERT_TRUE((M2_Pos_M - 5.0) <= 15.0, 'residu 14,75 m -> aucun depassement de butee');
END_TEST
